// TIA Portal project "11_End_LAGER_Projekt_261019" (V17)

(* hardware
DEVICE "S7300/ET200M-Station_4"  S7-300 station
   slot 0: "Profilschiene_0"  Rail  6ES7 390-1***0-0AA0
   slot 1: "PS 307 5A_1"  PS 307 5A  6ES7 307-1EA01-0AA0
   slot 2: "PLC_WBS_Bus"  CPU 314C-2 DP  6ES7 314-6CH04-0AB0  V3.3
      slot 0: "MPI-Schnittstelle_1"  MPI
      slot 1: "DP-Schnittstelle_1"  DP
      slot 2: "DI 24/DO 16_1"  DI24/DO16
      slot 3: "AI 5/AO 2_1"  AI5/AO2
      slot 4: "Zählen_1"  Counter
      slot 5: "Positionieren_1"  Positioning
   slot 4: "DI 64x24VDC sinking/souring_1"  DI64 x 24VDC  6ES7 321-1BP00-0AA0
   slot 5: "DI 64x24VDC sinking/souring_2"  DI64 x 24VDC  6ES7 321-1BP00-0AA0
   slot 6: "DI 64x24VDC sinking/souring_3"  DI64 x 24VDC  6ES7 321-1BP00-0AA0
   slot 7: "DI 64x24VDC sinking/souring_4"  DI64 x 24VDC  6ES7 321-1BP00-0AA0
   slot 8: "DO 64x24VDC/0.3A sourcing_1"  DO64 x 24VDC / 0.3A, P  6ES7 322-1BP00-0AA0
   slot 9: "DO 64x24VDC/0.3A sourcing_2"  DO64 x 24VDC / 0.3A, P  6ES7 322-1BP00-0AA0
   slot 10: "DO 64x24VDC/0.3A sourcing_3"  DO64 x 24VDC / 0.3A, P  6ES7 322-1BP00-0AA0
   slot 11: "DO 64x24VDC/0.3A sourcing_4"  DO64 x 24VDC / 0.3A, P  6ES7 322-1BP00-0AA0
DEVICE "PC-System_1"  SIMATIC PC station
   slot 0: "SIMATIC PC-Station"  Rail  SIMATIC PC-Station  V1.0
      slot 125: "Stationmanager"  Station_Manager  V6.0.4
   slot 1: "HMI_RT_1"  WinCC RT Advanced  6AV2 104-0xxxx-xxxx  17.0.0.0
      slot 33792: "Computerschnittstelle"  Host interface
   slot 3: "CP 5711_1"  CP 5711  6GK1 571-1AA00  V7.1.1
*)

// ===== PLC "PLC_WBS_Bus"  CPU 314C-2 DP =====

VAR_GLOBAL   // PLC tag table "Standard-Variablentabelle"
   "test_taster" AT %M26.1 : Bool;
   "Tag_1" AT %M100.1 : Bool;
END_VAR

VAR_GLOBAL   // PLC tag table "Betriebsart"
   "S0_HS" AT %E0.0 : Bool;   // Hauptschalter 0-Aus, 1-Ein
   "S1_Not_Halt" AT %E0.1 : Bool;   // Not-Halt NC
   "S2_START" AT %E0.2 : Bool;   // Taster START NO
   "S3_STOP" AT %E0.3 : Bool;   // Taster STOP NC
   "Res_E06" AT %E0.6 : Bool;
   "Res_E07" AT %E0.7 : Bool;
   "Res_E10" AT %E1.0 : Bool;
   "Res_E11" AT %E1.1 : Bool;
   "Res_E12" AT %E1.2 : Bool;
   "Res_E13" AT %E1.3 : Bool;
   "Res_E14" AT %E1.4 : Bool;
   "Res_E15" AT %E1.5 : Bool;
   "Res_E16" AT %E1.6 : Bool;
   "Factory_IO_RUN" AT %E1.7 : Bool;   // Rückmeldung Factory IO läuft
   "P1_MS_RT" AT %A0.0 : Bool;   // Meldesäule Rot
   "P2_MS_GE" AT %A0.1 : Bool;   // Meldesäule Gelb
   "P3_MS_GN" AT %A0.2 : Bool;   // Meldesäule Grün
   "P10_START" AT %A0.3 : Bool;   // Anzeige grün in START-Taster
   "P11_STOP" AT %A0.4 : Bool;   // Anzeige gelb in START-Taster
   "Res_A0.5" AT %A0.5 : Bool;
   "P12_Anfahrwarnung" AT %A0.6 : Bool;   // Rundumleuchte System
   "P13_Sirene" AT %A0.7 : Bool;   // Sirene System
   "Res_A12" AT %A1.2 : Bool;
   "Res_A13" AT %A1.3 : Bool;
   "Res_A14" AT %A1.4 : Bool;
   "Res_A15" AT %A1.5 : Bool;
   "Res_A16" AT %A1.6 : Bool;
   "Res_A17" AT %A1.7 : Bool;
   "Log_1" AT %M0.1 : Bool;   // statisch "1"
   "Log_0" AT %M0.0 : Bool;   // statisch "0"
   "Takt_1HZ" AT %M100.5 : Bool;   // Taktmerker 1 Hz
   "Anzeige_Anzahl_Teile_BL" AT %AW22 : Int;   // Anzeige Teile blau im Lager
   "Anzeige_Anzahl_Teile_GN" AT %AW24 : Int;   // Anzeige Teile grün im Lager
   "Start_Merker" AT %M26.0 : Bool;
   "S4_Auswahl_GN" AT %E0.4 : Bool;   // Taster Auswahl Teile grün NO
   "S5_Auswahl_BL" AT %E0.5 : Bool;   // Taster Auswahl Teile blau NO
   "P14_Auswahl_GN" AT %A1.0 : Bool;   // Anzeige Auswahl grün Taster
   "P15_Auswahl_BL" AT %A1.1 : Bool;   // Anzeige Auswahl blau Taster
   "M_False" AT %M202.0 : Bool;
   "M_True" AT %M202.1 : Bool;
   "Takt_2,5Hz" AT %M100.2 : Bool;
   "Pult_EW" AT %EW0 : Word;
   "Pult_AW" AT %AW0 : Word;
END_VAR

VAR_GLOBAL   // PLC tag table "Lager"
   "B8001_RB8001" AT %E2.0 : Bool;   // Transportband-Anfang
   "B8802_RB8001" AT %E2.1 : Bool;   // Transportband-Ende
   "B8003_RB8002" AT %E2.2 : Bool;   // Transportband-Anfang
   "B8004_RB8002" AT %E2.3 : Bool;   // Transportband-Ende
   "B8005_RB8003" AT %E2.4 : Bool;   // Transportband-Anfang
   "B8006_RB8003" AT %E2.5 : Bool;   // Transportband-Ende
   "B8007_OT_BL" AT %E2.6 : Bool;
   "B8008_OT_GN" AT %E2.7 : Bool;
   "B8020_STAPL_8001_Endlage_links" AT %E3.0 : Bool;   // Regaltransportgerät
   "B8021_STAPL_8001_Mittel_Pos" AT %E3.1 : Bool;   // Regaltransportgerät
   "B8022_STAPL_8001_Endlage_rechts" AT %E3.2 : Bool;   // Regaltransportgerät
   "B8023_STAPL_Bew_X_aktiv" AT %E3.3 : Bool;   // Regaltransportgerät
   "B8024_STAPL_Bew_Z_aktiv" AT %E3.4 : Bool;   // Regaltransportgerät
   "Res_E35" AT %E3.5 : Bool;
   "Res_E36" AT %E3.6 : Bool;
   "Res_E37" AT %E3.7 : Bool;
   "RB8001" AT %A2.0 : Bool;
   "RB8002" AT %A2.1 : Bool;
   "RB8003" AT %A2.2 : Bool;
   "STAPL_8001_Palette_heben" AT %A2.3 : Bool;
   "STAPL_8001_links_ausfahren" AT %A2.4 : Bool;
   "STAPL_8001_rechts_ausfahren" AT %A2.5 : Bool;
   "P8001_Warnung_Bewegung_1" AT %A2.6 : Bool;   // Rundumleuchte
   "P8002_Warnung_Bewegung_2" AT %A2.7 : Bool;   // Rundumleuchte
   "Res_A30" AT %A3.0 : Bool;
   "Res_A31" AT %A3.1 : Bool;
   "Res_A32" AT %A3.2 : Bool;
   "Res_A33" AT %A3.3 : Bool;
   "Res_A34" AT %A3.4 : Bool;
   "Res_A35" AT %A3.5 : Bool;
   "Res_A36" AT %A3.6 : Bool;
   "Emitter_1" AT %A3.7 : Bool;   // Emitter_1
   "STAPL_8001_Fachposition" AT %AW20 : Int;
END_VAR

VAR_GLOBAL   // PLC tag table "Versand_1"
   "B9001_RB9001" AT %E4.0 : Bool;   // Transportband-Anfang
   "B9002_RB9001" AT %E4.1 : Bool;   // Transportband-Ende
   "B9003_RB9002" AT %E4.2 : Bool;   // Transportband-Anfang
   "B9004_RB9002" AT %E4.3 : Bool;   // Transportband-Ende
   "B9005_RB9003" AT %E4.4 : Bool;   // Transportband-Anfang
   "B9006_RB9003" AT %E4.5 : Bool;   // Transportband-Ende
   "B9007_OT_BL" AT %E4.6 : Bool;   // Farberkennung blau
   "B9008_OT_GN" AT %E4.7 : Bool;   // Farberkennung grün
   "B9020_STAPL_9001_Endlage_links" AT %E5.0 : Bool;   // Regaltransportgerät
   "B9021_STAPL_9001_Mittel_Pos" AT %E5.1 : Bool;   // Regaltransportgerät
   "B9022_STAPL_9001_Endlage_rechts" AT %E5.2 : Bool;   // Regaltransportgerät
   "B9023_STAPL_Bew_X_aktiv" AT %E5.3 : Bool;   // Regaltransportgerät
   "B9024_STAPL_Bew_Z_aktiv" AT %E5.4 : Bool;   // Regaltransportgerät
   "RB9001" AT %A4.0 : Bool;
   "RB9002" AT %A4.1 : Bool;
   "RB9003" AT %A4.2 : Bool;
   "STAPL_9001_Palette_heben" AT %A4.3 : Bool;
   "STAPL_9001_links_ausfahren" AT %A4.4 : Bool;
   "STAPL_9001_rechts_ausfahren" AT %A4.5 : Bool;
   "P9001_Warnung_Bewegung_1" AT %A4.6 : Bool;   // Rundumleuchte
   "P9002_Warnung_Bewegung_2" AT %A4.7 : Bool;   // Rundumleuchte
   "Res_A37" AT %A5.7 : Bool;
   "STAPL_9001_Fachposition" AT %AW26 : Int;
END_VAR

TYPE "Datenspeicher"
   STRUCT
      DatumUhrzeit : Date_And_Time;
      Materialfarbe : String[10];
      Materialfarbe_Nummer : Int;
      Frei : Bool := TRUE;
   END_STRUCT;
END_TYPE

TYPE "Pult_Output"
   STRUCT
      P1_MS_RT : Bool;
      P2_MS_GE : Bool;
      P3_MS_GN : Bool;
      P10_START : Bool;
      P11_STOP : Bool;
      "Res_A0.5" : Bool;
      P12_Anfahrwarnung : Bool;
      P13_Sirene : Bool;
      P14_Auswahl_GN : Bool;
      P15_Auswahl_BL : Bool;
      Res_A12 : Bool;
      Res_A13 : Bool;
      Res_A14 : Bool;
      Res_A15 : Bool;
      Res_A16 : Bool;
      Res_A17 : Bool;
   END_STRUCT;
END_TYPE

TYPE "Datenaustausch_Lager"
   STRUCT
      Anlage_Ein : Bool;
      Anlage_Betriebsbereit : Bool;
      Anlage_Stop : Bool;
      NotHalt : Bool;
      Position : Int;
   END_STRUCT;
END_TYPE

TYPE "Datenaustausch_Versand"
   STRUCT
      Anlage_Ein : Bool;
      Anlage_Betriebsbereit : Bool;
      Anlage_Stop : Bool;
      NotHalt : Bool;
      i_Blau : Bool;
      i_Grün : Bool;
      i_630_Grundstellung : Bool;
      i_640_RB_Frei : Bool;
      i_fehler : Bool;
      i_Blau_Anzahl : Int;
      i_Grün_Anzahl : Int;
      Position : Int;
   END_STRUCT;
END_TYPE

TYPE "Pult_Input"
   STRUCT
      S0_HS : Bool;
      S1_Not_Halt : Bool;
      S2_START : Bool;
      S3_STOP : Bool;
      S4_Auswahl_GN : Bool;
      S5_Auswahl_BL : Bool;
      Res_E06 : Bool;
      Res_E07 : Bool;
      Res_E10 : Bool;
      Res_E11 : Bool;
      Res_E12 : Bool;
      Res_E13 : Bool;
      Res_E14 : Bool;
      Res_E15 : Bool;
      Res_E16 : Bool;
      Factory_IO_RUN : Bool;
   END_STRUCT;
END_TYPE

// folder: LAGER/DB

DATA_BLOCK "HochregallagerDB"   // DB1
{ S7_Optimized_Access := 'FALSE' }
VERSION : 0.1
   VAR
      Freigabe : Bool := False;   // Freigabe der Anlage
      Palette_Bereit_Pos55 : Bool := True;   // Palette an Übergabeposition 55 zur Übernahme bereit
      Stapler_Fachposition_Eingabe : Int := 1;   // Zielposition des Staplers: 1–54 Lagerfach, 55 Übergabe
      Stapler_Auftrag_Aktiv : Bool;   // Stapler bearbeitet einen Auftrag
      Stapler_Auftrag_Fertig : Bool;   // Staplerauftrag abgeschlossen
      Stapler_Stoerung : Bool;   // Störung am Stapler vorhanden
      Farbe : Int;   // Erkannter Farbcode: 1 = Blau, 2 = Grün, 4 = Fehler
      Stappler_Aktuele_Farbe : Int;   // Farbcode der aktuell vom Stapler transportierten Palette
      Automatik : Bool := True;   // Automatikbetrieb aktiviert
      Motors_Ein : Bool;   // Einschaltsignal für die Rollenbahnmotoren
      Neue_Palette : Bool;   // Signal für eine neue Palette
      HMI_X_Bewegung : Int;   // Horizontale Position für die Stapleranimation im HMI
      HMI_Z_Bewegung : Int;   // Vertikale Position für die Stapleranimation im HMI
      Reset_Counter : Bool;   // Zähler zurücksetzen
      Lagerplaetze : Array[1..54] of "Datenspeicher";   // Lagerdaten der 54 Lagerplätze: Belegung, Farbe und Einlagerungszeit
      Anzahl_Blau : Int;   // Anzahl der eingelagerten blauen Paletten
      Anzahl_Gruen : Int;   // Anzahl der eingelagerten grünen Paletten
      Anzahl_Unbekannte_Farbe : Int;   // Anzahl der eingelagerten Unbekannte Paletten
      Einlagerungsposition : Int;   // Nummer des Lagerplatzes für die zu speichernden Palettendaten (1–54)
      Stapler_In_Bewegung : Bool;   // Stacker in motion
      Rollenbahn_In_Bewegung : Bool;   // Conveyor in motion
      Stoerung_Aktiv : Bool;   // Eine Störung liegt vor.
      Warnung_Aktiv : Bool;   // Eine Warnung liegt vor.
      Warnung_Wenig_Freie_Plaetze : Bool;   // TRUE: Warnschwelle erreicht oder unterschritten; auch bei vollem Lager aktiv.
      Lager_Voll : Bool;   // TRUE: Alle Lagerplaetze sind belegt.
      Stopp_Am_Zyklusende : Bool;
   END_VAR
BEGIN
END_DATA_BLOCK

DATA_BLOCK "HMI_Eingaben_DB"   // DB8
{ S7_Optimized_Access := 'FALSE' }
VERSION : 0.1
   VAR
      HMI_Start : Bool;
      HMI_Stop : Bool := TRUE;
      HMI_Not_Halt : Bool := TRUE;
      HMI_Hauptschalter : Bool;
      HMI_Start_Anzeige : Bool;
   END_VAR
BEGIN
END_DATA_BLOCK

// folder: LAGER/Instance

DATA_BLOCK "FB_Paketempfang_Rollenbahn_DB"   // DB2
{ S7_Optimized_Access := 'FALSE' }
VERSION : 0.1
// stored: InstanceOfName FB_Paketempfang_Rollenbahn
"FB_Paketempfang_Rollenbahn"
BEGIN
END_DATA_BLOCK

DATA_BLOCK "FB_Stapler_Ablauf_DB"   // DB3
{ S7_Optimized_Access := 'FALSE' }
VERSION : 0.1
// stored: InstanceOfName FB_Stapler_Ablauf
"FB_Stapler_Ablauf"
BEGIN
END_DATA_BLOCK

DATA_BLOCK "FB_Lagerverwaltung_DB"   // DB4
{ S7_Optimized_Access := 'FALSE' }
VERSION : 0.1
// stored: InstanceOfName FB_Lagerverwaltung
"FB_Lagerverwaltung"
BEGIN
END_DATA_BLOCK

DATA_BLOCK "FB_ControlPanel_DB"   // DB7
{ S7_Optimized_Access := 'FALSE' }
VERSION : 0.1
// stored: InstanceOfName FB_ControlPanel
"FB_ControlPanel"
BEGIN
END_DATA_BLOCK

DATA_BLOCK "Lager_Aufrufen_DB"   // DB9
{ S7_Optimized_Access := 'FALSE' }
VERSION : 0.1
// stored: InstanceOfName Lager_Aufrufen
"Lager_Aufrufen"
BEGIN
END_DATA_BLOCK

// folder: LAGER/Lager_AWL

DATA_BLOCK "Lager_Daten"   // DB8000
{ S7_Optimized_Access := 'FALSE' }
VERSION : 0.1
   VAR
      Lagerfach : Array[1..54] of Int;   // 1 = blau, 2 = grün, 0 = leer
   END_VAR
BEGIN
   Lagerfach[1] := 1;
   Lagerfach[2] := 2;
   Lagerfach[3] := 1;
   Lagerfach[4] := 2;
   Lagerfach[5] := 2;
   Lagerfach[6] := 2;
   Lagerfach[7] := 2;
   Lagerfach[8] := 2;
   Lagerfach[9] := 2;
   Lagerfach[10] := 2;
   Lagerfach[11] := 1;
   Lagerfach[12] := 1;
   Lagerfach[54] := 1;
   Lagerfach[13] := 1;
   Lagerfach[14] := 1;
   Lagerfach[15] := 1;
   Lagerfach[16] := 1;
   Lagerfach[17] := 1;
   Lagerfach[18] := 2;
   Lagerfach[19] := 2;
   Lagerfach[20] := 1;
   Lagerfach[21] := 2;
   Lagerfach[22] := 2;
   Lagerfach[23] := 2;
   Lagerfach[24] := 2;
   Lagerfach[25] := 2;
   Lagerfach[26] := 2;
   Lagerfach[27] := 2;
   Lagerfach[28] := 2;
   Lagerfach[29] := 1;
   Lagerfach[30] := 1;
   Lagerfach[31] := 1;
   Lagerfach[32] := 1;
   Lagerfach[33] := 1;
   Lagerfach[34] := 1;
   Lagerfach[35] := 1;
   Lagerfach[36] := 1;
   Lagerfach[37] := 1;
   Lagerfach[38] := 1;
   Lagerfach[39] := 2;
   Lagerfach[40] := 2;
   Lagerfach[41] := 2;
   Lagerfach[42] := 1;
   Lagerfach[43] := 1;
   Lagerfach[44] := 1;
   Lagerfach[45] := 1;
   Lagerfach[46] := 2;
   Lagerfach[47] := 2;
   Lagerfach[48] := 2;
   Lagerfach[49] := 2;
   Lagerfach[50] := 2;
   Lagerfach[51] := 0;
   Lagerfach[52] := 2;
   Lagerfach[53] := 1;
END_DATA_BLOCK

// folder: Versand

DATA_BLOCK "600_Versand_Main_DB"   // DB10
{ S7_Optimized_Access := 'FALSE' }
AUTHOR : DJonas
VERSION : 0.1
// stored: InstanceOfName 600_Versand_Main
"600_Versand_Main"
BEGIN
END_DATA_BLOCK

// folder: (top level)

ORGANIZATION_BLOCK "Main"   // OB1, FBD
TITLE = "Main Program Sweep (Cycle)"
{ S7_Optimized_Access := 'FALSE' }
VERSION : 0.1
   VAR_TEMP
      OB1_EV_CLASS : Byte;   // Bits 0-3 = 1 (Coming event), Bits 4-7 = 1 (Event class 1)
      OB1_SCAN_1 : Byte;   // 1 (Cold restart scan 1 of OB 1), 3 (Scan 2-n of OB 1)
      OB1_PRIORITY : Byte;   // Priority of OB Execution
      OB1_OB_NUMBR : Byte;   // 1 (Organization block 1, OB1)
      OB1_RESERVED_1 : Byte;   // Reserved for system
      OB1_RESERVED_2 : Byte;   // Reserved for system
      OB1_PREV_CYCLE : Int;   // Cycle time of previous OB1 scan (milliseconds)
      OB1_MIN_CYCLE : Int;   // Minimum cycle time of OB1 (milliseconds)
      OB1_MAX_CYCLE : Int;   // Maximum cycle time of OB1 (milliseconds)
      OB1_DATE_TIME : Date_And_Time;   // Date and time OB1 started
   END_VAR
BEGIN

REGION Network 1
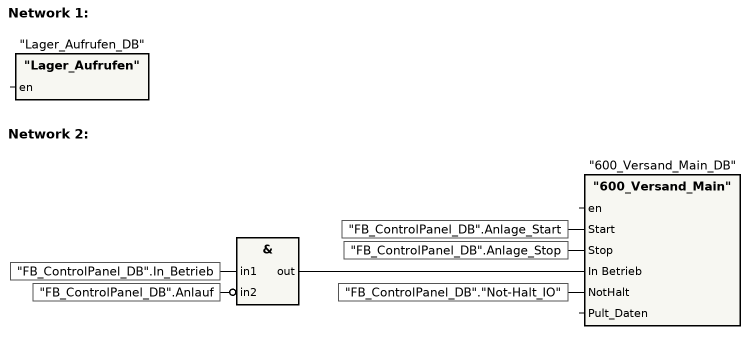
   "Lager_Aufrufen_DB"();   // "Lager_Aufrufen"
END_REGION

REGION Network 2
   "600_Versand_Main_DB"(Start := "FB_ControlPanel_DB".Anlage_Start,   // "600_Versand_Main"
                         Stop := "FB_ControlPanel_DB".Anlage_Stop,
                         "In Betrieb" := "FB_ControlPanel_DB".In_Betrieb AND NOT "FB_ControlPanel_DB".Anlauf,
                         NotHalt := "FB_ControlPanel_DB"."Not-Halt_IO");
END_REGION
END_ORGANIZATION_BLOCK

// folder: LAGER

FUNCTION_BLOCK "Lager_Aufrufen"   // FB4, FBD
{ S7_Optimized_Access := 'FALSE' }
VERSION : 0.1
BEGIN

REGION Network 1: Bedienpanel Signale verarbeiten
   // Start-, Stopp- und Not-Halt-Signale von Bedienpanel und HMI zusammenführen und an den FB_ControlPanel übergeben. Hauptschalter, Factory-I/O-Betriebsstatus und Palettenanzahlen einlesen sowie Meldeleuchten ansteuern.
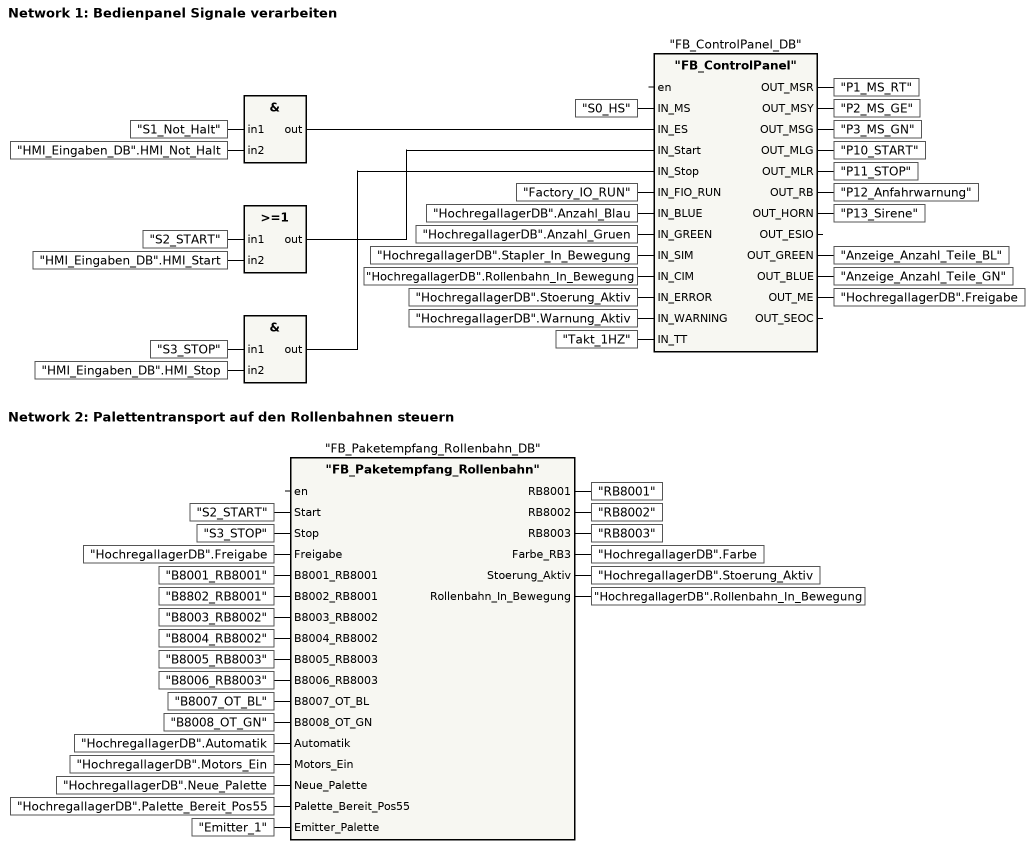
   "FB_ControlPanel_DB"(IN_MS := "S0_HS",   // "FB_ControlPanel"
                        IN_ES := "S1_Not_Halt" AND "HMI_Eingaben_DB".HMI_Not_Halt,
                        IN_Start := "S2_START" OR "HMI_Eingaben_DB".HMI_Start,
                        IN_Stop := "S3_STOP" AND "HMI_Eingaben_DB".HMI_Stop,
                        IN_FIO_RUN := "Factory_IO_RUN",
                        IN_BLUE := "HochregallagerDB".Anzahl_Blau,
                        IN_GREEN := "HochregallagerDB".Anzahl_Gruen,
                        IN_SIM := "HochregallagerDB".Stapler_In_Bewegung,
                        IN_CIM := "HochregallagerDB".Rollenbahn_In_Bewegung,
                        IN_ERROR := "HochregallagerDB".Stoerung_Aktiv,
                        IN_WARNING := "HochregallagerDB".Warnung_Aktiv,
                        IN_TT := "Takt_1HZ",
                        OUT_MSR => "P1_MS_RT",
                        OUT_MSY => "P2_MS_GE",
                        OUT_MSG => "P3_MS_GN",
                        OUT_MLG => "P10_START",
                        OUT_MLR => "P11_STOP",
                        OUT_RB => "P12_Anfahrwarnung",
                        OUT_HORN => "P13_Sirene",
                        OUT_GREEN => "Anzeige_Anzahl_Teile_BL",
                        OUT_BLUE => "Anzeige_Anzahl_Teile_GN",
                        OUT_ME => "HochregallagerDB".Freigabe);
END_REGION

REGION Network 2: Palettentransport auf den Rollenbahnen steuern
   // FB_Paketempfang_Rollenbahn aufrufen, Sensorsignale und Farberkennung auswerten sowie die drei Rollenbahnen abhängig von Start, Stopp und Freigabe ansteuern.
   "FB_Paketempfang_Rollenbahn_DB"(Start := "S2_START",   // "FB_Paketempfang_Rollenbahn"
                           Stop := "S3_STOP",
                           Freigabe := "HochregallagerDB".Freigabe,
                           B8001_RB8001 := "B8001_RB8001",
                           B8002_RB8001 := "B8802_RB8001",
                           B8003_RB8002 := "B8003_RB8002",
                           B8004_RB8002 := "B8004_RB8002",
                           B8005_RB8003 := "B8005_RB8003",
                           B8006_RB8003 := "B8006_RB8003",
                           B8007_OT_BL := "B8007_OT_BL",
                           B8008_OT_GN := "B8008_OT_GN",
                           Automatik := "HochregallagerDB".Automatik,
                           Motors_Ein := "HochregallagerDB".Motors_Ein,
                           Neue_Palette := "HochregallagerDB".Neue_Palette,
                           Palette_Bereit_Pos55 := "HochregallagerDB".Palette_Bereit_Pos55,
                           Emitter_Palette := "Emitter_1",
                           RB8001 => "RB8001",
                           RB8002 => "RB8002",
                           RB8003 => "RB8003",
                           Farbe_RB3 => "HochregallagerDB".Farbe,
                           Stoerung_Aktiv => "HochregallagerDB".Stoerung_Aktiv,
                           Rollenbahn_In_Bewegung => "HochregallagerDB".Rollenbahn_In_Bewegung);
END_REGION

REGION Network 3: Staplerablauf steuern
   // Der Baustein verarbeitet Freigabe, Stopp und Sensorsignale, steuert die Palettenaufnahme und Einlagerung und meldet den Auftragsstatus.
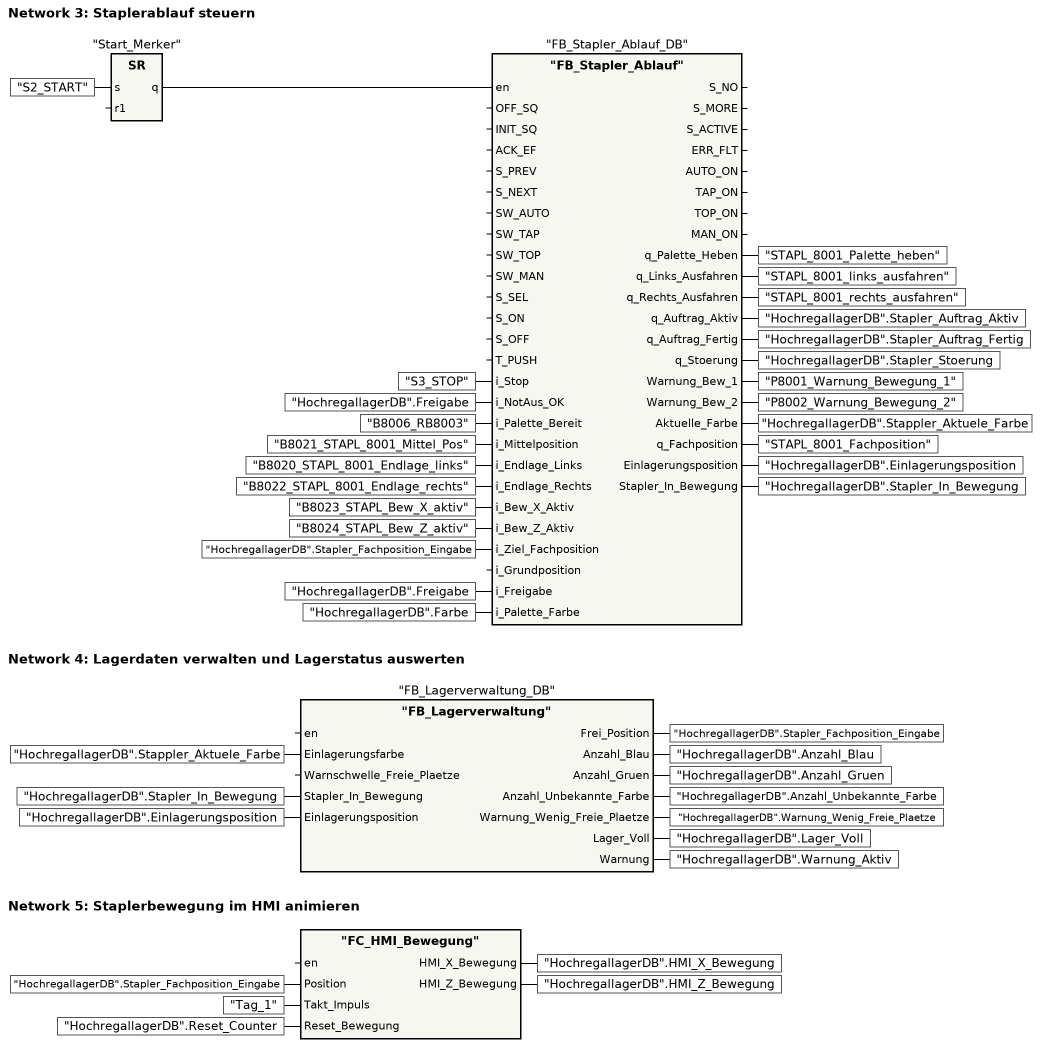
   IF "S2_START" THEN
       "Start_Merker" := TRUE;   // SR flip-flop
   END_IF;
   IF "Start_Merker" THEN
       "FB_Stapler_Ablauf_DB"(i_Stop := "S3_STOP",   // "FB_Stapler_Ablauf"
                              i_NotAus_OK := "HochregallagerDB".Freigabe,
                              i_Palette_Bereit := "B8006_RB8003",
                              i_Mittelposition := "B8021_STAPL_8001_Mittel_Pos",
                              i_Endlage_Links := "B8020_STAPL_8001_Endlage_links",
                              i_Endlage_Rechts := "B8022_STAPL_8001_Endlage_rechts",
                              i_Bew_X_Aktiv := "B8023_STAPL_Bew_X_aktiv",
                              i_Bew_Z_Aktiv := "B8024_STAPL_Bew_Z_aktiv",
                              i_Ziel_Fachposition := "HochregallagerDB".Stapler_Fachposition_Eingabe,
                              i_Freigabe := "HochregallagerDB".Freigabe,
                              i_Palette_Farbe := "HochregallagerDB".Farbe,
                              q_Palette_Heben => "STAPL_8001_Palette_heben",
                              q_Links_Ausfahren => "STAPL_8001_links_ausfahren",
                              q_Rechts_Ausfahren => "STAPL_8001_rechts_ausfahren",
                              q_Auftrag_Aktiv => "HochregallagerDB".Stapler_Auftrag_Aktiv,
                              q_Auftrag_Fertig => "HochregallagerDB".Stapler_Auftrag_Fertig,
                              q_Stoerung => "HochregallagerDB".Stapler_Stoerung,
                              Warnung_Bew_1 => "P8001_Warnung_Bewegung_1",
                              Warnung_Bew_2 => "P8002_Warnung_Bewegung_2",
                              Aktuelle_Farbe => "HochregallagerDB".Stappler_Aktuele_Farbe,
                              q_Fachposition => "STAPL_8001_Fachposition",
                              Einlagerungsposition => "HochregallagerDB".Einlagerungsposition,
                              Stapler_In_Bewegung => "HochregallagerDB".Stapler_In_Bewegung);
   END_IF;
END_REGION

REGION Network 4: Lagerdaten verwalten und Lagerstatus auswerten
   // FB_Lagerverwaltung aufrufen, Palettendaten speichern und freie Lagerplätze ermitteln. Paletten nach Farbe zählen und Warnungen bei wenigen freien Plätzen oder vollem Lager ausgeben.
   "FB_Lagerverwaltung_DB"(Einlagerungsfarbe := "HochregallagerDB".Stappler_Aktuele_Farbe,   // "FB_Lagerverwaltung"
                           Stapler_In_Bewegung := "HochregallagerDB".Stapler_In_Bewegung,
                           Einlagerungsposition := "HochregallagerDB".Einlagerungsposition,
                           Frei_Position => "HochregallagerDB".Stapler_Fachposition_Eingabe,
                           Anzahl_Blau => "HochregallagerDB".Anzahl_Blau,
                           Anzahl_Gruen => "HochregallagerDB".Anzahl_Gruen,
                           Anzahl_Unbekannte_Farbe => "HochregallagerDB".Anzahl_Unbekannte_Farbe,
                           Warnung_Wenig_Freie_Plaetze => "HochregallagerDB".Warnung_Wenig_Freie_Plaetze,
                           Lager_Voll => "HochregallagerDB".Lager_Voll,
                           Warnung => "HochregallagerDB".Warnung_Aktiv);
END_REGION

REGION Network 5: Staplerbewegung im HMI animieren
   // FC_HMI_Bewegung aufrufen, um aus der Fachposition und dem Taktsignal die X- und Z-Verschiebung für die HMI-Animation zu berechnen.
   "FC_HMI_Bewegung"(Position := "HochregallagerDB".Stapler_Fachposition_Eingabe,
                     Takt_Impuls := "Tag_1",
                     Reset_Bewegung := "HochregallagerDB".Reset_Counter,
                     HMI_X_Bewegung => "HochregallagerDB".HMI_X_Bewegung,
                     HMI_Z_Bewegung => "HochregallagerDB".HMI_Z_Bewegung);
END_REGION
END_FUNCTION_BLOCK

// folder: LAGER/FB

FUNCTION_BLOCK "FB_Paketempfang_Rollenbahn"   // FB1, FBD
TITLE = Paketempfang und Rollenbahnsteuerung
{ S7_Optimized_Access := 'FALSE' }
VERSION : 0.1
// - Der FB übernimmt die Steuerung des Palettentransports vom Emitter bis zur Übergabeposition 55 des Regalstapelsystems.
   VAR_INPUT
      Start : Bool;   // Anlage/Funktion freigegeben
      Stop : Bool;   // Stop-Anforderung
      Freigabe : Bool;   // Freigabe für Paketempfang und Rollenbahnsteuerung
      B8001_RB8001 : Bool;   // Sensor Palette auf Rollenbahn 1
      B8002_RB8001 : Bool;   // Sensor Ende Rollenbahn 1
      B8003_RB8002 : Bool;   // Sensor Palette auf Rollenbahn 2
      B8004_RB8002 : Bool;   // Sensor Ende Rollenbahn 2
      B8005_RB8003 : Bool;   // Sensor Palette auf Rollenbahn 3
      B8006_RB8003 : Bool;   // Sensor Ende Rollenbahn 3 (Palette hat Position 55 erreicht)
      B8007_OT_BL : Bool;   // optischer Sensor erkennt Blau
      B8008_OT_GN : Bool;   // optischer Sensor erkennt Grün
      Automatik : Bool;   // Betriebsart Automatik
      Motors_Ein : Bool;
      Neue_Palette : Bool;
   END_VAR
   VAR_OUTPUT
      RB8001 : Bool;   // Motor Rollenbahn 1
      RB8002 : Bool;   // Motor Rollenbahn 2
      RB8003 : Bool;   // Motor Rollenbahn 3
      Farbe_RB3 : Int;   // (1: Blau / 2:Grün / 4:Fehler)
      Stoerung_Aktiv : Bool;
      Rollenbahn_In_Bewegung : Bool;
   END_VAR
   VAR_IN_OUT
      Palette_Bereit_Pos55 : Bool;   // Palette steht zur Übernahme bereit
      Emitter_Palette : Bool;   // Emitter hat eine Palette bereitgestellt
   END_VAR
   VAR
      Empfang_Aktiv : Bool;   // FB bearbeitet aktuell eine Palette
      Betriebsfreigabe : Bool;   // Gespeicherte Freigabe für den Betrieb der Rollenbahnsteuerung
      Start_P_Merker : Bool;   // Flankenmerker für positive Flanke des Startsignals
      Emitter_P_Merker : Bool;   // Flankenmerker für positive Flanke des Emitter-Signals
      S2_N_Merker : Bool;   // Flankenmerker für negative Flanke von Sensor B8002
      S2_P_Merker : Bool;   // Merker für die positieve Flanke von Sensor 2
      S3_P_Merker : Bool;   // Flankenmerker für positive Flanke von Sensor B8003
      S4_N_Merker : Bool;   // Flankenmerker für negative Flanke von Sensor B8004
      S5_P_Merker : Bool;   // Flankenmerker für positive Flanke von Sensor B8005
      S6_N_Merker : Bool;   // Merker für die negative Flanke von Sensor 6
      S6_P_Merker : Bool;   // Flankenmerker für positive Flanke von Sensor B8006
      RB1_Merker : Bool;   // Speichermerker für Ansteuerung Rollenbahn 1
      RB2_Merker : Bool;   // Speichermerker für Ansteuerung Rollenbahn 2
      S3_N_Merker : Bool;
      RB3_Merker : Bool;   // Speichermerker für Ansteuerung Rollenbahn 3
      SBL_P_Merker : Bool;   // Flankenmerker für positive Flanke des Sensors Blau
      SGR_P_Merker : Bool;   // Flankenmerker für positive Flanke des Sensors Grün
      Palette_auf_RB1 : Bool;   // Palette befindet sich auf Rollenbahn 1
      Palette_auf_RB2 : Bool;   // Palette befindet sich auf Rollenbahn 2
      Palette_auf_RB3 : Bool;   // Palette befindet sich auf Rollenbahn 3
      Farbe_RB2 : Int;   // Erkannte Palettenfarbe auf Rollenbahn RB8002
      IEC_Timer_0_Instance : TON;   // Instanz des TON-Timers für Laufzeitüberwachung
      IEC_Timer_0_Instance_1 : TON;   // TON-Timerinstanz für Zeitüberwachung
      s_warnung_1 : Bool;   // Rollenbahn länger als zulässige Zeit aktiv
      s_warnung_2 : Bool;   // Sensor B8003_RB8002 länger als zulässige Zeit aktiv
      s_warnung_3 : Bool;
      IEC_Timer_0_Instance_2 : TON;
      Farbe_Merker : Bool;
      IEC_Timer_0_Instance_3 : TON;
   END_VAR
   VAR_TEMP   // added for the SCL form of the ladder/FBD networks
      _w1 : Bool;
      _w2 : Bool;
      _w3 : Bool;
      _w4 : Bool;
   END_VAR
BEGIN

REGION Network 1: Betriebsfreigabe
   // - Betriebsfreigabe über Start setzen und bei Stop bzw. fehlender Freigabe zurücksetzen.
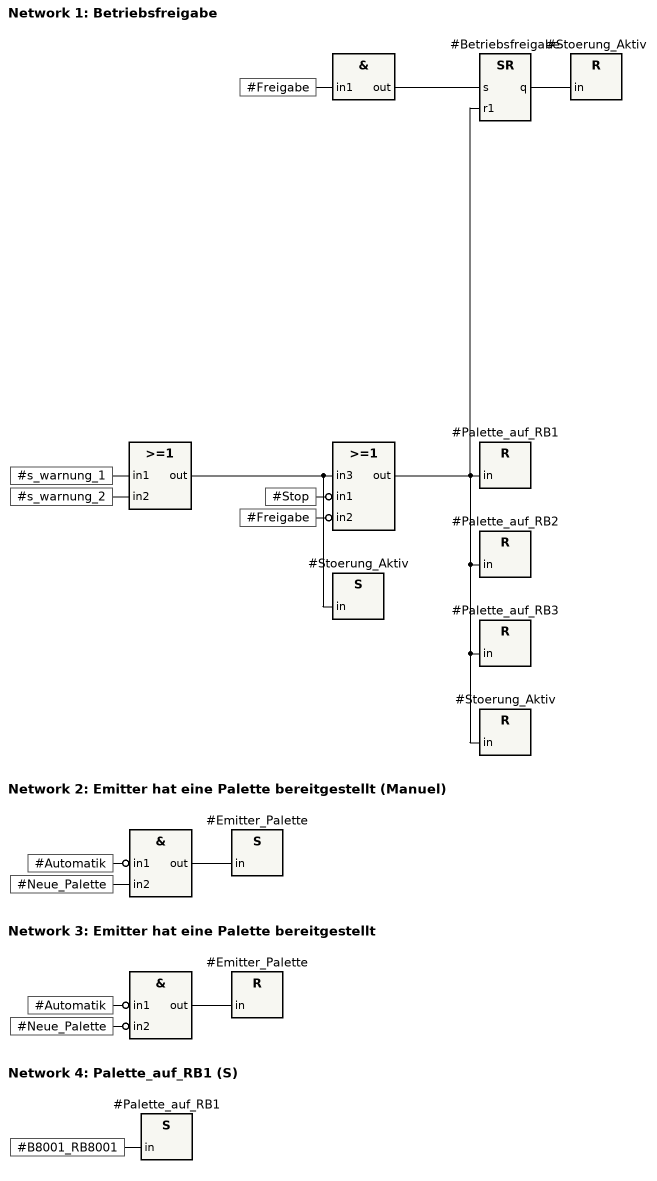
   #_w1 := #s_warnung_1 OR #s_warnung_2;
   #_w2 := #_w1 OR NOT #Stop OR NOT #Freigabe;
   IF #Freigabe THEN
       #Betriebsfreigabe := TRUE;   // SR flip-flop
   END_IF;
   IF #_w2 THEN #Betriebsfreigabe := FALSE; END_IF;
   IF #Betriebsfreigabe THEN #Stoerung_Aktiv := FALSE; END_IF;
   IF #_w2 THEN
       #Palette_auf_RB1 := FALSE;
       #Palette_auf_RB2 := FALSE;
       #Palette_auf_RB3 := FALSE;
       #Stoerung_Aktiv := FALSE;
   END_IF;
   IF #_w1 THEN #Stoerung_Aktiv := TRUE; END_IF;
END_REGION

REGION Network 2: Emitter hat eine Palette bereitgestellt (Manuel)
   IF NOT #Automatik AND #Neue_Palette THEN #Emitter_Palette := TRUE; END_IF;
END_REGION

REGION Network 3: Emitter hat eine Palette bereitgestellt
   IF NOT #Automatik AND NOT #Neue_Palette THEN #Emitter_Palette := FALSE; END_IF;
END_REGION

REGION Network 4: Palette_auf_RB1 (S)
   IF #B8001_RB8001 THEN #Palette_auf_RB1 := TRUE; END_IF;
END_REGION

REGION Network 5: Motor Rollenbahn 1
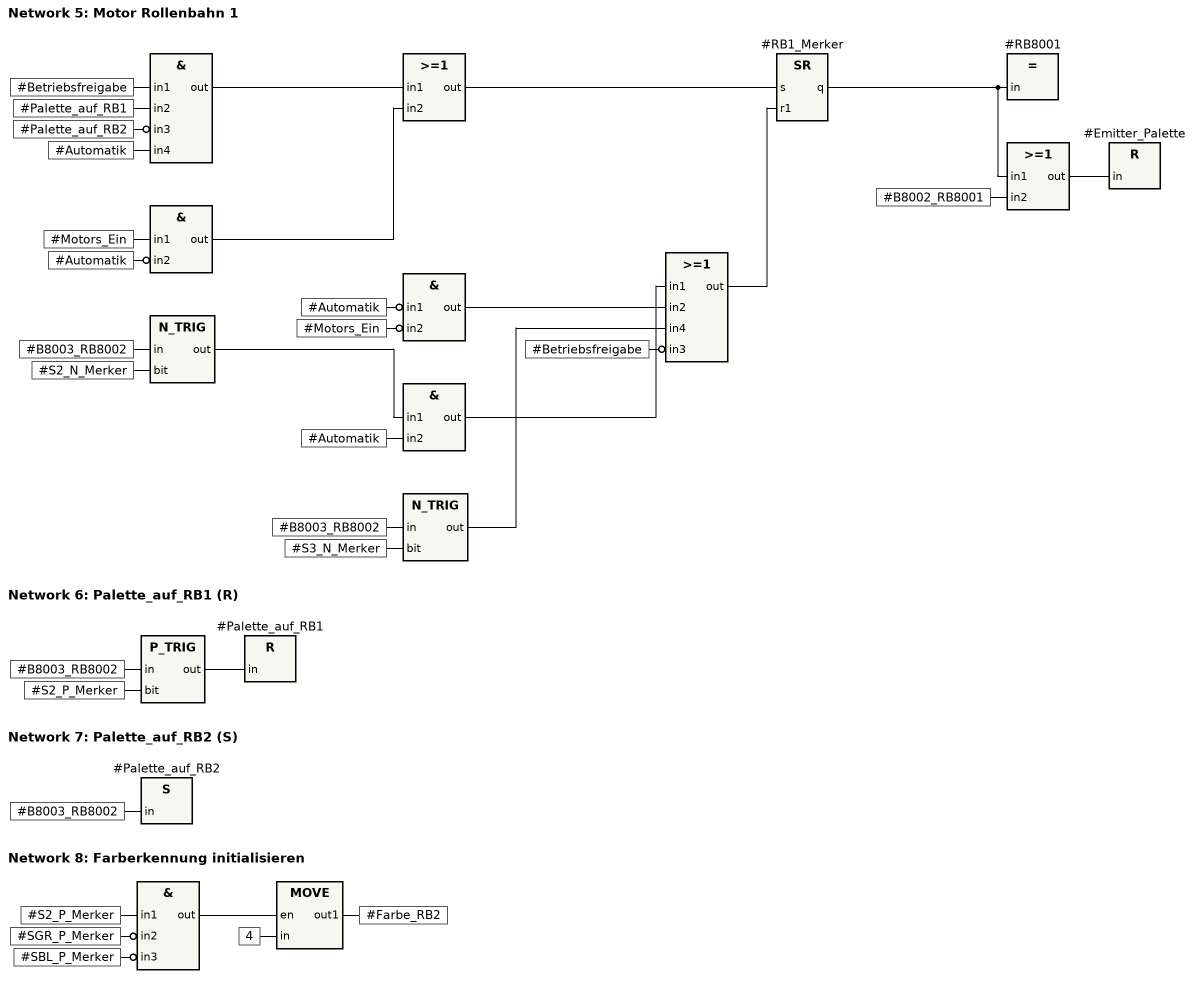
   #_w1 := NOT #B8003_RB8002 AND #S2_N_Merker;   // falling edge
   #S2_N_Merker := #B8003_RB8002;
   #_w2 := NOT #B8003_RB8002 AND #S3_N_Merker;   // falling edge
   #S3_N_Merker := #B8003_RB8002;
   IF (#Betriebsfreigabe AND #Palette_auf_RB1 AND NOT #Palette_auf_RB2 AND #Automatik) OR (#Motors_Ein AND NOT #Automatik) THEN
       #RB1_Merker := TRUE;   // SR flip-flop
   END_IF;
   IF (#_w1 AND #Automatik) OR (NOT #Automatik AND NOT #Motors_Ein) OR #_w2 OR NOT #Betriebsfreigabe THEN
       #RB1_Merker := FALSE;
   END_IF;
   #RB8001 := #RB1_Merker;
   IF #RB1_Merker OR #B8002_RB8001 THEN #Emitter_Palette := FALSE; END_IF;
END_REGION

REGION Network 6: Palette_auf_RB1 (R)
   #_w1 := #B8003_RB8002 AND NOT #S2_P_Merker;   // rising edge
   #S2_P_Merker := #B8003_RB8002;
   IF #_w1 THEN #Palette_auf_RB1 := FALSE; END_IF;
END_REGION

REGION Network 7: Palette_auf_RB2 (S)
   IF #B8003_RB8002 THEN #Palette_auf_RB2 := TRUE; END_IF;
END_REGION

REGION Network 8: Farberkennung initialisieren
   IF #S2_P_Merker AND NOT #SGR_P_Merker AND NOT #SBL_P_Merker THEN #Farbe_RB2 := 4; END_IF;
END_REGION

REGION Network 9: Motor Rollenbahn 2 / Farberkennung (Blau,Grün)
   // (1: Blau / 2:Grün / 4:Fehler)
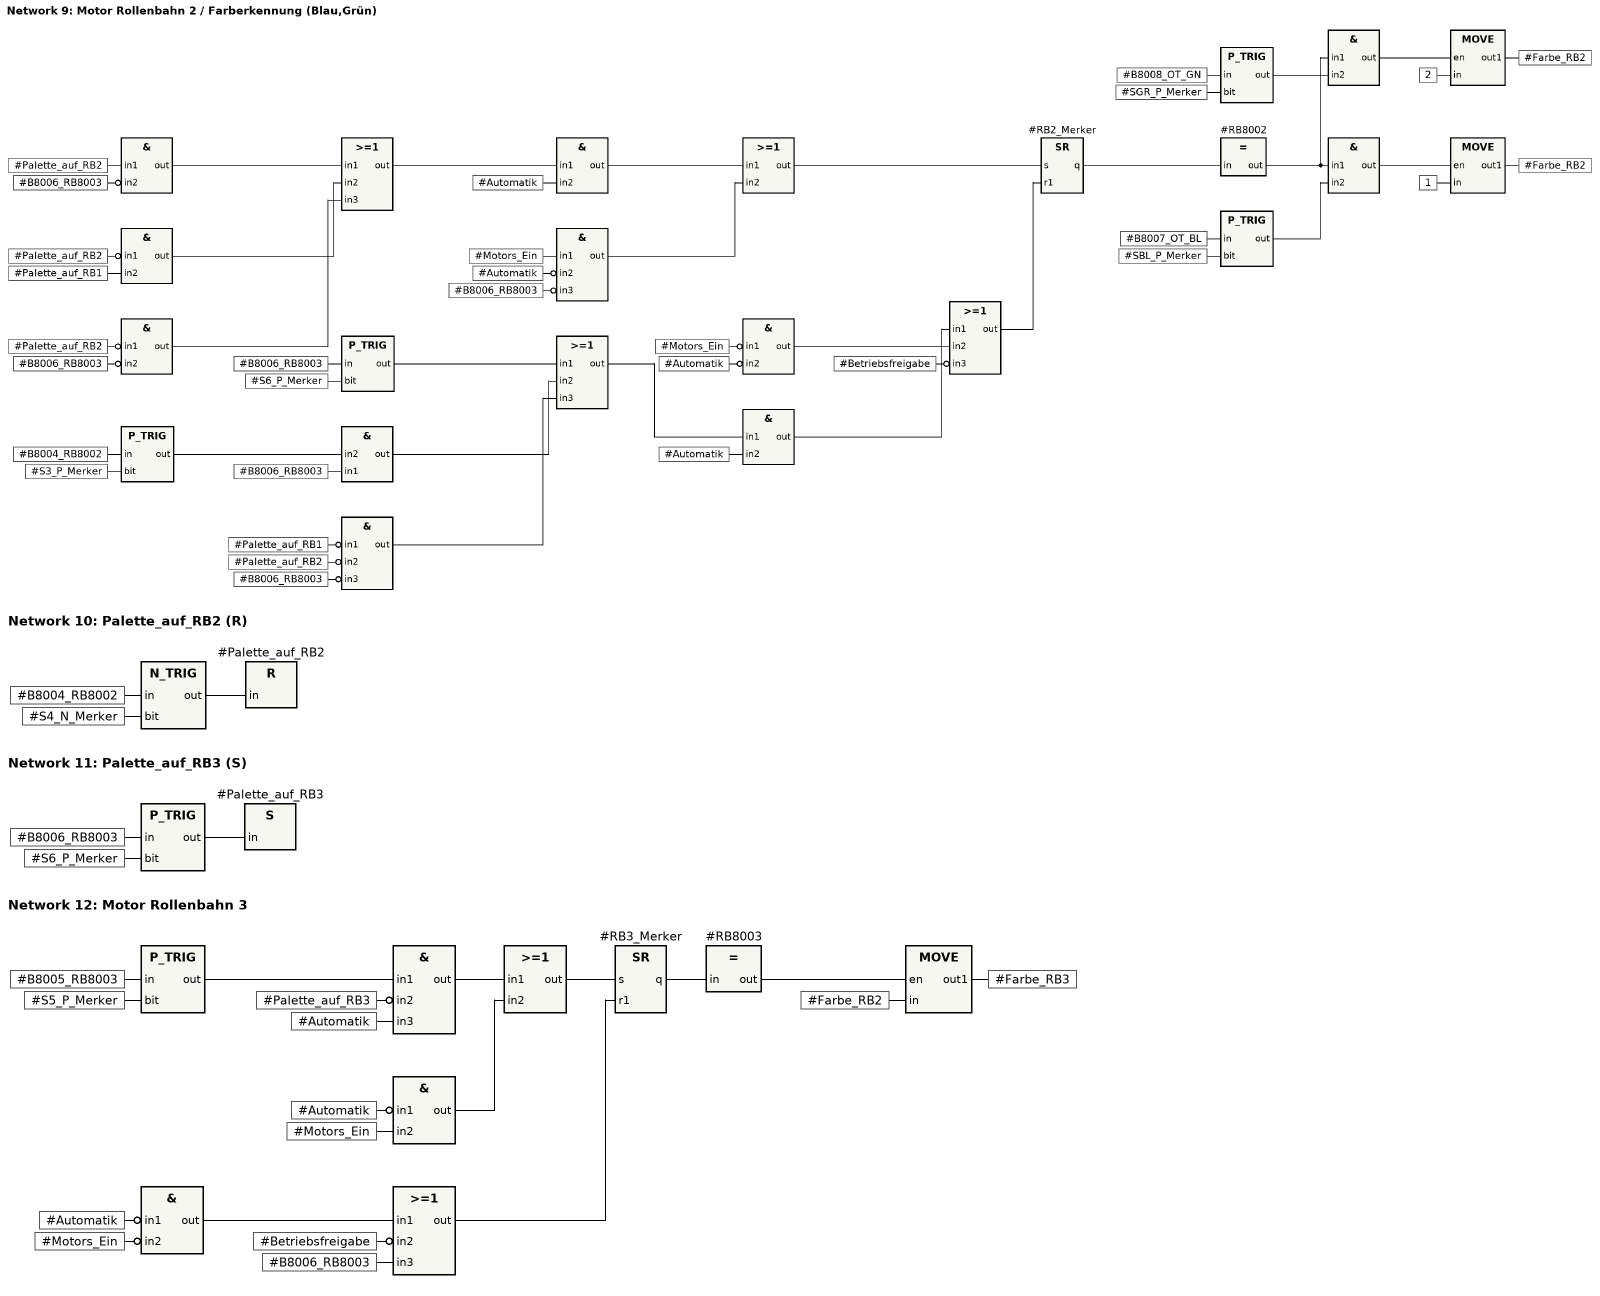
   #_w1 := #B8006_RB8003 AND NOT #S6_P_Merker;   // rising edge
   #S6_P_Merker := #B8006_RB8003;
   #_w2 := #B8004_RB8002 AND NOT #S3_P_Merker;   // rising edge
   #S3_P_Merker := #B8004_RB8002;
   IF (((#Palette_auf_RB2 AND NOT #B8006_RB8003) OR (NOT #Palette_auf_RB2 AND #Palette_auf_RB1) OR (NOT #Palette_auf_RB2 AND NOT #B8006_RB8003)) AND #Automatik) OR (#Motors_Ein AND NOT #Automatik AND NOT #B8006_RB8003) THEN
       #RB2_Merker := TRUE;   // SR flip-flop
   END_IF;
   IF ((#_w1 OR (#_w2 AND #B8006_RB8003) OR (NOT #Palette_auf_RB1 AND NOT #Palette_auf_RB2 AND NOT #B8006_RB8003)) AND #Automatik) OR (NOT #Motors_Ein AND NOT #Automatik) OR NOT #Betriebsfreigabe THEN
       #RB2_Merker := FALSE;
   END_IF;
   #RB8002 := #RB2_Merker;
   #_w3 := #B8008_OT_GN AND NOT #SGR_P_Merker;   // rising edge
   #SGR_P_Merker := #B8008_OT_GN;
   IF #RB2_Merker AND #_w3 THEN #Farbe_RB2 := 2; END_IF;
   #_w4 := #B8007_OT_BL AND NOT #SBL_P_Merker;   // rising edge
   #SBL_P_Merker := #B8007_OT_BL;
   IF #RB2_Merker AND #_w4 THEN #Farbe_RB2 := 1; END_IF;
END_REGION

REGION Network 10: Palette_auf_RB2 (R)
   #_w1 := NOT #B8004_RB8002 AND #S4_N_Merker;   // falling edge
   #S4_N_Merker := #B8004_RB8002;
   IF #_w1 THEN #Palette_auf_RB2 := FALSE; END_IF;
END_REGION

REGION Network 11: Palette_auf_RB3 (S)
   #_w1 := #B8006_RB8003 AND NOT #S6_P_Merker;   // rising edge
   #S6_P_Merker := #B8006_RB8003;
   IF #_w1 THEN #Palette_auf_RB3 := TRUE; END_IF;
END_REGION

REGION Network 12: Motor Rollenbahn 3
   // Farbe_RB3 (1: Blau / 2:Grün)
   #_w1 := #B8005_RB8003 AND NOT #S5_P_Merker;   // rising edge
   #S5_P_Merker := #B8005_RB8003;
   IF (#_w1 AND NOT #Palette_auf_RB3 AND #Automatik) OR (NOT #Automatik AND #Motors_Ein) THEN
       #RB3_Merker := TRUE;   // SR flip-flop
   END_IF;
   IF (NOT #Automatik AND NOT #Motors_Ein) OR NOT #Betriebsfreigabe OR #B8006_RB8003 THEN
       #RB3_Merker := FALSE;
   END_IF;
   #RB8003 := #RB3_Merker;
   IF #RB3_Merker THEN #Farbe_RB3 := #Farbe_RB2; END_IF;
END_REGION

REGION Network 13: Palette_auf_RB3 (R)
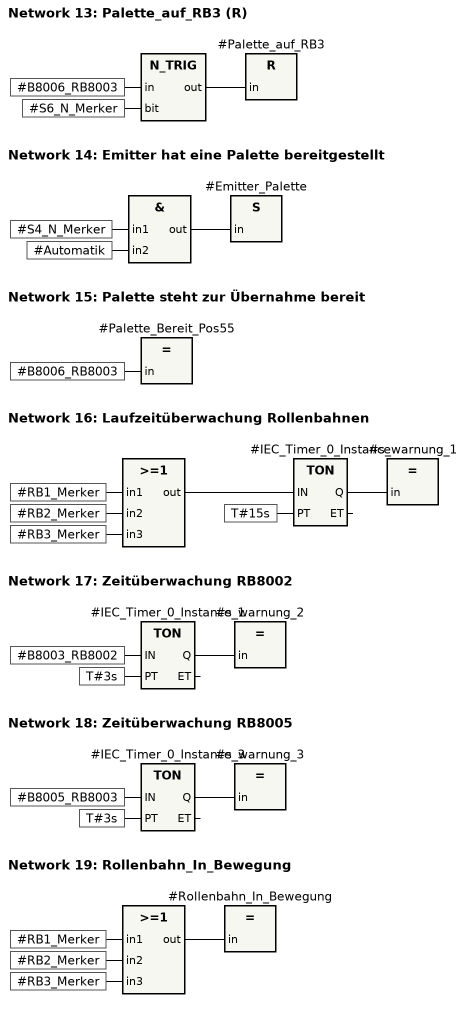
   #_w1 := NOT #B8006_RB8003 AND #S6_N_Merker;   // falling edge
   #S6_N_Merker := #B8006_RB8003;
   IF #_w1 THEN #Palette_auf_RB3 := FALSE; END_IF;
END_REGION

REGION Network 14: Emitter hat eine Palette bereitgestellt
   IF #S4_N_Merker AND #Automatik THEN #Emitter_Palette := TRUE; END_IF;
END_REGION

REGION Network 15: Palette steht zur Übernahme bereit
   #Palette_Bereit_Pos55 := #B8006_RB8003;
END_REGION

REGION Network 16: Laufzeitüberwachung Rollenbahnen
   // 14-s-Zeitüberwachung für aktive Rollenbahn. Bei Zeitüberschreitung wird s_warnung_1 gesetzt.
   #IEC_Timer_0_Instance.TON(IN := #RB1_Merker OR #RB2_Merker OR #RB3_Merker, PT := T#15s);
   #s_warnung_1 := #IEC_Timer_0_Instance.Q;
END_REGION

REGION Network 17: Zeitüberwachung RB8002
   // Ist der Sensor B8003_RB8002 länger als 4 s aktiv, wird die Warnung s_warnung_2 gesetzt.
   #IEC_Timer_0_Instance_1.TON(IN := #B8003_RB8002, PT := T#3s);
   #s_warnung_2 := #IEC_Timer_0_Instance_1.Q;
END_REGION

REGION Network 18: Zeitüberwachung RB8005
   #IEC_Timer_0_Instance_3.TON(IN := #B8005_RB8003, PT := T#3s);
   #s_warnung_3 := #IEC_Timer_0_Instance_3.Q;
END_REGION

REGION Network 19: Rollenbahn_In_Bewegung
   #Rollenbahn_In_Bewegung := #RB1_Merker OR #RB2_Merker OR #RB3_Merker;
END_REGION
END_FUNCTION_BLOCK

FUNCTION_BLOCK "FB_Stapler_Ablauf"   // FB2, GRAPH
{ S7_Optimized_Access := 'FALSE' }
VERSION : 0.1
   VAR_INPUT
      OFF_SQ : Bool := false;   // Kette ausschalten
      INIT_SQ : Bool := false;   // Kette in Initialzustand versetzen
      ACK_EF : Bool := false;   // Alle Fehler und Störungen quittieren
      S_PREV : Bool := false;   // Vorherigen Schritt am Parameter S_NO ausgeben
      S_NEXT : Bool := false;   // Nächsten Schritt am Parameter S_NO anzeigen
      SW_AUTO : Bool := false;   // Automatischer Betrieb
      SW_TAP : Bool := false;   // Halbautomatisch/Weiterschalten mit Transition
      SW_TOP : Bool := false;   // Halbautomatisch/Ignoriere Transition
      SW_MAN : Bool := false;   // Handbetrieb
      S_SEL : Int := 0;   // Schritt auswählen, der an S_NO ausgegeben werden soll
      S_ON : Bool := false;   // Schritt aktivieren, der an Parameter S_NO anliegt
      S_OFF : Bool := false;   // Schritt deaktivieren, der an Parameter S_NO anliegt
      T_PUSH : Bool := false;   // Schaltfreigabe für Transition im halbautomatischen Betrieb
      i_Stop : Bool;
      i_NotAus_OK : Bool;   // TRUE = kein Not-Aus / Anlage sicher
      i_Palette_Bereit : Bool;   // Palette wartet auf Einlagerung
      i_Mittelposition : Bool;   // Gabel in Mittelposition
      i_Endlage_Links : Bool;   // Gabel links vollständig ausgefahren
      i_Endlage_Rechts : Bool;   // Gabel rechts vollständig ausgefahren
      i_Bew_X_Aktiv : Bool;   // X-Bewegung aktiv
      i_Bew_Z_Aktiv : Bool;   // Z-Bewegung aktiv
      i_Ziel_Fachposition : Int;   // Zielposition für die Einlagerung
      i_Grundposition : Int := 55;   // Grundposition, bei dir 55
      i_Freigabe : Bool;
      i_Palette_Farbe : Int;   // (1: Blau / 2:Grün / 4:Fehler)
   END_VAR
   VAR_OUTPUT
      S_NO : Int := 0;   // Schrittnummer
      S_MORE : Bool := false;   // Weitere Schritte sind vorhanden und können in S_NO angezeigt werden.
      S_ACTIVE : Bool := false;   // Schritt, der an Parameter S_NO angezeigt wird, ist aktiv
      ERR_FLT : Bool := false;   // Sammelfehler Interlock oder Supervision
      AUTO_ON : Bool := false;   // Automatischer Betrieb eingeschaltet
      TAP_ON : Bool := false;   // Halbautomatischer Betrieb/Schritt mit Transition eingeschaltet
      TOP_ON : Bool := false;   // Halbautomatischer Betrieb/Ignoriere Transition eingeschaltet
      MAN_ON : Bool := false;   // Handbetrieb eingeschaltet
      q_Palette_Heben : Bool;   // Gabel links ausfahren
      q_Links_Ausfahren : Bool;   // Gabel links ausfahren
      q_Rechts_Ausfahren : Bool;   // Gabel rechts ausfahren
      q_Auftrag_Aktiv : Bool;   // Einlagerungsauftrag läuft
      q_Auftrag_Fertig : Bool;   // Auftrag abgeschlossen
      q_Stoerung : Bool;   // Störung im Staplerablauf
      Warnung_Bew_1 : Bool;
      Warnung_Bew_2 : Bool;
      Aktuelle_Farbe : Int;   // (1: Blau / 2:Grün / 4:Fehler)
      q_Fachposition : Int;   // Sollposition des Staplers
      Einlagerungsposition : Int;
      Stapler_In_Bewegung : Bool;
   END_VAR
   VAR
      SWITCH : Array[0..0] of DWord;
      SW_SQTS : Array[0..12] of Byte;
      SW_ADDR : Word := 16#1A;
      G7T_0 : GraphTransition;
      G7S_0 : GraphStep;
      PRE_CRIT : Array[0..0] of DWord;
      POST_CRIT : Array[0..0] of DWord;
      TVX : Array[0..2] of Byte;
      TTX : Array[0..2] of Byte;
      TSX : Array[0..2] of Byte;
      S00X : Array[0..2] of Byte;
      SOFFX : Array[0..2] of Byte;
      SONX : Array[0..2] of Byte;
      SAX : Array[0..2] of Byte;
      SERRX : Array[0..13] of Byte;
      SMX : Array[0..13] of Byte;
      S0X : Array[0..13] of Byte;
      S1X : Array[0..13] of Byte;
      S_DISPLAY : Int;   // Interne Anzeige des Ausgangsparameters S_NO
      S_SEL_OLD : Int;   // Vorheriger Wert an S_SEL
      S_DISPIDX : Byte;   // Index des Schritts, der an S_NO anliegt
      T_DISPIDX : Byte;   // Index der Transition, die an T_NO anliegt
      MOPEDGE : Struct
         AUTO : Bool := false;
         MAN : Bool := false;
         TAP : Bool := false;
         TOP : Bool := false;
         ACK_S : Bool := false;
         REG_S : Bool := false;
         T_PREV : Bool := false;
         T_NEXT : Bool := false;
         LOCK : Bool := false;
         SUP : Bool := false;
         ACKREQ : Bool := false;
         SSKIP : Bool := false;
         OFF : Bool := false;
         INIT : Bool := false;
         HALT : Bool := false;
         TMS_HALT : Bool := false;
         OPS_ZERO : Bool := false;
         SACT_DISP : Bool := false;
         SEF_DISP : Bool := false;
         SALL_DISP : Bool := false;
         S_PREV : Bool := false;
         S_NEXT : Bool := false;
         S_SELOK : Bool := false;
         S_ON : Bool := false;
         S_OFF : Bool := false;
         T_PUSH : Bool := false;
         REG : Bool := false;
         ACK : Bool := false;
         IL_PERM : Bool := false;
         T_PERM : Bool := false;
         ILP_MAN : Bool := false;
      END_STRUCT;
      MOP : Struct   // Betriebsart
         AUTO : Bool := true;   // Zustand: Automatischer Betrieb
         MAN : Bool := false;   // Zustand: Handbetrieb
         TAP : Bool := false;   // Zustand: Halbautomatisch/Weiterschalten mit Transition
         TOP : Bool := false;   // Zustand: Halbautomatisch/Ignoriere Transition
         ACK_S : Bool := false;   // Anforderung: Schritt quittieren, der an Parameter S_NO anliegt
         REG_S : Bool := false;   // Anforderung: Schritt registrieren, der an Parameter S_NO anliegt
         T_PREV : Bool := false;   // Anforderung: Vorherige gültige Transition am Parameter T_NO ausgeben
         T_NEXT : Bool := false;   // Anforderung: Nächste gültige Transition am Parameter T_NO ausgeben
         LOCK : Bool := true;   // Zustand: Interlockbearbeitung aktiviert
         SUP : Bool := true;   // Zustand: Supervisionsbearbeitung aktiviert
         ACKREQ : Bool := true;   // Zustand: Quittierung erforderlich
         SSKIP : Bool := false;   // Zustand: "Schritte überspringen" aktiviert
         OFF : Bool := false;   // Anforderung: Alle Schritte deaktivieren
         INIT : Bool := true;   // Anforderung: Kette in Initialzustand schalten
         HALT : Bool := false;   // Zustand: Kette schaltet nicht weiter
         TMS_HALT : Bool := false;   // Zustand: Alle internen Zeiten angehalten
         OPS_ZERO : Bool := false;   // Zustand: Alle mit N, L, D bearbeitete Operanden auf 0 gesetzt
         SACT_DISP : Bool := true;   // Zustand: Nur aktive Schritte anzeigen
         SEF_DISP : Bool := false;   // Zustand: Nur fehlerhafte und gestörte Schritte anzeigen
         SALL_DISP : Bool := false;   // Zustand: Alle Schritte anzeigen
         S_PREV : Bool := false;   // Anforderung: Vorherigen Schritt am Parameter S_NO ausgeben
         S_NEXT : Bool := false;   // Anforderung: Nächsten Schritt am Parameter S_NO ausgeben
         S_SELOK : Bool := false;   // Anforderung: Schrittnummer, die am Parameter S_SEL anliegt, am Parameter S_NO ausgeben
         S_ON : Bool := false;   // Anforderung: Schritt aktivieren, der am Parameter S_NO anliegt
         S_OFF : Bool := false;   // Anforderung: Schritt deaktivieren, der am Parameter S_NO anliegt
         T_PUSH : Bool := false;   // Anforderung: Schaltfreigabe für Transition
         REG : Bool := false;   // Anforderung: Alle Interlock- und Supervisionsfehler registrieren
         ACK : Bool := false;   // Anforderung: Alle Interlock- und Supervisionsfehler quittieren
         IL_PERM : Bool := false;   // Zustand: Permanente Bearbeitung aller Interlocks
         T_PERM : Bool := false;   // Zustand: Permanente Bearbeitung aller Transitionen
         ILP_MAN : Bool := false;   // Zustand: Permanente Bearbeitung aller Interlocks im Handbetrieb
      END_STRUCT;
      TICKS : Struct   // Zeittakte
         DELTA : Time := T#0ms;   // Zeitdifferenz zwischen zwei Zyklen
         OLD : Time := T#0ms;   // 10 ms Taktzählerstand im letzten Zyklus
         NEW : Time := T#0ms;   // 10 ms Taktzählerstand in diesem Zyklus
      END_STRUCT;
      SQ_FLAGS : Struct   // Kettenmerker
         ERR_FLT : Bool := false;   // Sammelfehler Interlock und Supervision
         ERROR : Bool := false;   // Sammelfehler Interlock
         FAULT : Bool := false;   // Sammelfehler Supervision
         RT_FAIL : Bool := false;   // Laufzeitfehler
         NO_SNO : Bool := false;   // Angeforderte Schrittnummer nicht gefunden
         NF_OFL : Bool := false;   // Überlauf: Zu viele Anforderungen ON oder OFF
         SA_OFL : Bool := false;   // Überlauf: Zu viele Schritte aktiv
         TV_OFL : Bool := false;   // Überlauf: Zu viele gültige Transitionen
         MSG_OFL : Bool := false;   // Überlauf: Nicht genügend Systemressourcen fü ALARM_S
         NO_SWI : Bool := false;   // Nicht Schalten in diesem Zyklus
         CYC_OP : Bool := false;   // Zyklische Bearbeitung der Kette nach Initialisierung
         AS_MSG : Bool := false;   // Meldungen zur Laufzeit durch Anweisung aktiviert oder deaktiviert
         AS_SEND : Bool := false;   // Meldungen von WR_USMSG senden oder nur in Diagnosepuffer eintragen
         SQ_BUSY : Bool := false;   // Interner Flankenmerker für Vorgangsbearbeitung
         SA_BUSY : Bool := false;   // Interner Flankenmerker für Vorgangsbearbeitung
         AS_SIG : Bool := false;   // Flankenmerker für Meldungen von Alarm_S und Alarm_SQ
      END_STRUCT;
      S_PTR : DWord := 16#7F0;
      S_PTR2 : DWord := 16#0;
      S_PTR3 : DWord := 16#1760;
      S_PTR4 : DWord := 16#16F0;
      T_PTR : DWord := 16#1680;
      C_AR2 : DWord := 16#0;
      M_FBDB : DWord := 16#20000;
      M_SNO : Word := 16#0;
      M_EVID : Word := 16#0;
      M_EVIL : DWord;
      M_EVSV : DWord;
      M_EV : DWord := 16#15B0;
      CRIT : Array[0..31] of Bool;
      S_START : Byte := 16#0;
      S_IDX : Byte := 16#0;
      S_INT : Int := 72;
      S_TMP : Byte := 16#0;
      T_START : Byte := 16#0;
      T_IDX : Byte := 16#0;
      T_TMP : Byte := 16#0;
      T_TMP2 : Byte := 16#00;
      TV_POT : Byte := 16#0E;
      RETURN1 : Byte := 16#0;
      RETURN2 : Byte := 16#0;
      SINI : Array[0..2] of Byte;
      LSTT : Array[0..12] of Byte;
      ATAJ : Array[0..12] of Byte;
      ATAB : Array[0..12] of Byte;
      PSTT : Array[0..12] of Byte;
      NSTT : Array[0..12] of Byte;
      ASSJ : Array[0..12] of Byte;
      ASSB : Array[0..12] of Byte;
      PTTS : Array[0..12] of Byte;
      NTTS : Array[0..12] of Byte;
      PRE_CNT : Word := 16#1;
      POST_CNT : Word := 16#1;
      ADR_COND : Word := 16#0;
      MAX_TVAL : Byte := 16#1;
      MAX_SACT : Byte := 16#1;
      MAX_CRIT : Byte := 16#4;
      T_CNT : Byte := 16#C;
      SUP_CNT : Byte := 16#0;
      LOCK_CNT : Byte := 16#2;
      S_CNT : Byte := 16#C;
      SQ_CNT : Byte := 16#1;
      PRS_INPAR : DWord := 16#E000FEC8;
      PRS_OUTPAR : DWord := 16#E000800F;
      GC_FLAGS : Struct
         T_MACH : Byte := 16#EB;
         COND_ED : Byte := 16#E2;
         W_LEVEL : Byte := 16#D5;
         FB_IF : Byte := 16#FA;
         AS_MSG : Word := 16#0;
         SSB : Word := 16#108;
         DILG : Word := 16#3FC;
         ADDR_T0 : Word := 16#2E;
         CRIT_AVAIL : Bool := false;
         SSKIP_AVAIL : Bool := true;
         SSKIP_ON : Bool := false;
         ACK_REQ : Bool := true;
         SYNC_AVAIL : Bool := true;
         ILP_MAN : Bool := false;
         SWM_LOCKED : Bool := false;
         SAVE_SW : Bool := true;
      END_STRUCT;
      G7_FBMARK : Byte := 16#3C;
      G7_RELEASE : Byte := 16#3C;
      G7_ID2 : Byte := 16#37;
      G7_ID1 : Byte := 16#47;
   END_VAR
   // SW_SQTS[0] := 16#1;
   // TVX[0] := 16#1;
   // TTX[0] := 16#1;
   // TSX[0] := 16#1;
   // S00X[0] := 16#1;
   // SOFFX[0] := 16#1;
   // SONX[0] := 16#1;
   // SAX[0] := 16#1;
   // SERRX[0] := 16#1;
   // SMX[0] := 16#1;
   // S0X[0] := 16#1;
   // S1X[0] := 16#1;
   // SINI[0] := 16#2;
   // SINI[1] := 16#1;
   // SINI[2] := 0;
   // LSTT[0] := 0;
   // LSTT[1] := 0;
   // LSTT[2] := 0;
   // LSTT[3] := 0;
   // LSTT[4] := 0;
   // LSTT[5] := 0;
   // LSTT[6] := 0;
   // LSTT[7] := 0;
   // ATAJ[0] := 0;
   // ATAJ[1] := 16#1;
   // ATAJ[2] := 16#2;
   // ATAJ[3] := 16#3;
   // ATAJ[4] := 16#4;
   // ATAJ[5] := 16#5;
   // ATAJ[6] := 16#6;
   // ATAJ[7] := 16#7;
   // ATAB[0] := 0;
   // ATAB[1] := 16#1;
   // ATAB[2] := 16#2;
   // ATAB[3] := 16#3;
   // ATAB[4] := 16#4;
   // ATAB[5] := 16#5;
   // ATAB[6] := 16#6;
   // ATAB[7] := 16#7;
   // PSTT[0] := 0;
   // PSTT[1] := 16#1;
   // PSTT[2] := 16#2;
   // PSTT[3] := 16#3;
   // PSTT[4] := 16#4;
   // PSTT[5] := 16#5;
   // PSTT[6] := 16#6;
   // PSTT[7] := 16#7;
   // NSTT[0] := 16#1;
   // NSTT[1] := 16#2;
   // NSTT[2] := 16#3;
   // NSTT[3] := 16#4;
   // NSTT[4] := 16#5;
   // NSTT[5] := 16#6;
   // NSTT[6] := 16#7;
   // NSTT[7] := 16#8;
   // ASSJ[0] := 0;
   // ASSJ[1] := 16#1;
   // ASSJ[2] := 16#2;
   // ASSJ[3] := 16#3;
   // ASSJ[4] := 16#4;
   // ASSJ[5] := 16#5;
   // ASSJ[6] := 16#6;
   // ASSJ[7] := 16#7;
   // ASSB[0] := 0;
   // ASSB[1] := 16#1;
   // ASSB[2] := 16#2;
   // ASSB[3] := 16#3;
   // ASSB[4] := 16#4;
   // ASSB[5] := 16#5;
   // ASSB[6] := 16#6;
   // ASSB[7] := 16#7;
   // PTTS[0] := 0;
   // PTTS[2] := 16#1;
   // PTTS[3] := 16#2;
   // PTTS[4] := 16#3;
   // PTTS[5] := 16#4;
   // PTTS[6] := 16#5;
   // PTTS[7] := 16#6;
   // NTTS[0] := 0;
   // NTTS[1] := 16#1;
   // NTTS[2] := 16#2;
   // NTTS[3] := 16#3;
   // NTTS[4] := 16#4;
   // NTTS[5] := 16#5;
   // NTTS[6] := 16#6;
   // NTTS[7] := 16#7;
   // LSTT[8] := 0;
   // LSTT[9] := 0;
   // LSTT[10] := 0;
   // ATAJ[8] := 16#8;
   // ATAJ[9] := 16#9;
   // ATAJ[10] := 16#A;
   // ATAB[8] := 16#8;
   // ATAB[9] := 16#9;
   // ATAB[10] := 16#A;
   // PSTT[8] := 16#8;
   // PSTT[9] := 16#9;
   // PSTT[10] := 16#A;
   // NSTT[8] := 16#9;
   // NSTT[9] := 16#A;
   // NSTT[10] := 16#C;
   // ASSJ[8] := 16#8;
   // ASSJ[9] := 16#9;
   // ASSJ[10] := 16#A;
   // ASSB[8] := 16#8;
   // ASSB[9] := 16#9;
   // ASSB[10] := 16#A;
   // PTTS[8] := 16#7;
   // PTTS[9] := 16#8;
   // PTTS[10] := 16#9;
   // NTTS[8] := 16#8;
   // NTTS[9] := 16#9;
   // NTTS[10] := 16#A;
   // LSTT[11] := 16#1;
   // ATAJ[11] := 16#B;
   // ATAB[11] := 16#B;
   // PSTT[11] := 16#B;
   // NSTT[11] := 16#1;
   // ASSJ[11] := 16#B;
   // ASSB[11] := 16#B;
   // PTTS[11] := 16#C;
   // NTTS[11] := 16#B;
   // LSTT[12] := 0;
   // ATAJ[12] := 16#C;
   // ATAB[12] := 16#C;
   // PSTT[12] := 16#C;
   // NSTT[12] := 16#B;
   // ASSJ[12] := 16#C;
   // ASSB[12] := 16#C;
   // PTTS[12] := 16#A;
   // NTTS[12] := 16#C;
BEGIN
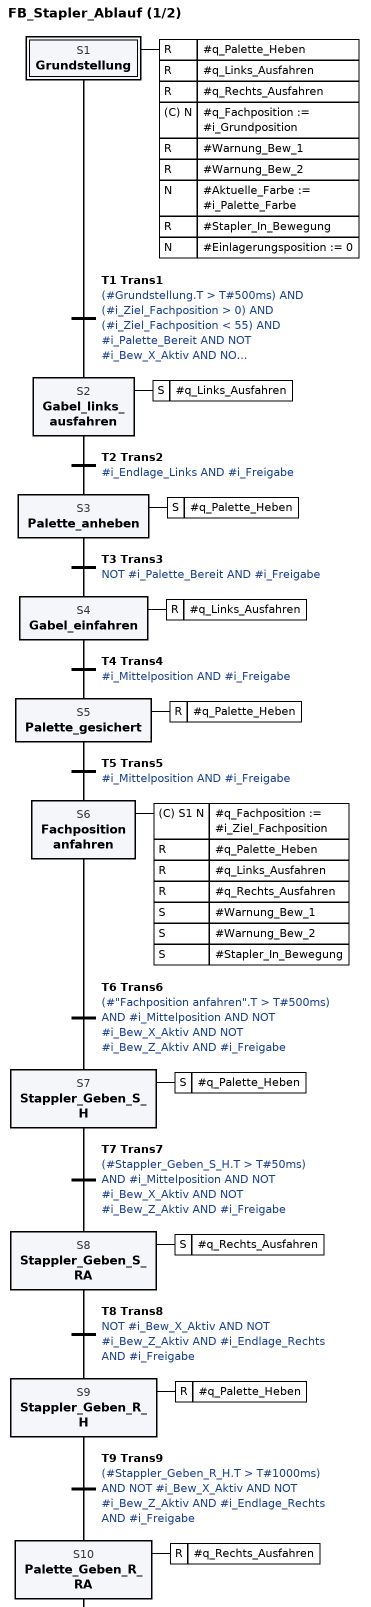
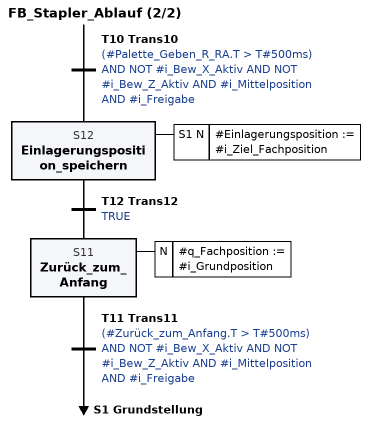
   // sequencer 1
   INITIAL_STEP Grundstellung:   // S1
      interlock C := #i_NotAus_OK AND #i_Stop;
      // - Stapler befindet sich in Grundstellung auf Position 55. Alle Ausgänge sind deaktiviert. Warten auf eine einlagerbereite Palette.
              R    #q_Palette_Heben
              R    #q_Links_Ausfahren
              R    #q_Rechts_Ausfahren
      (C)     N    #q_Fachposition := #i_Grundposition
              R    #Warnung_Bew_1
              R    #Warnung_Bew_2
              N    #Aktuelle_Farbe := #i_Palette_Farbe
              R    #Stapler_In_Bewegung
              N    #Einlagerungsposition := 0
   END_STEP
   TRANSITION Trans1 FROM Grundstellung TO Gabel_links_ausfahren   // T1
      := (#Grundstellung.T > T#500ms) AND (#i_Ziel_Fachposition > 0) AND (#i_Ziel_Fachposition < 55) AND #i_Palette_Bereit AND NOT #i_Bew_X_Aktiv AND NOT #i_Bew_Z_Aktiv AND #i_NotAus_OK AND #i_Stop AND #i_Freigabe;
   END_TRANSITION
   STEP Gabel_links_ausfahren:   // S2
              S    #q_Links_Ausfahren
   END_STEP
   TRANSITION Trans2 FROM Gabel_links_ausfahren TO Palette_anheben   // T2
      := #i_Endlage_Links AND #i_Freigabe;
   END_TRANSITION
   STEP Palette_anheben:   // S3
              S    #q_Palette_Heben
   END_STEP
   TRANSITION Trans3 FROM Palette_anheben TO Gabel_einfahren   // T3
      := NOT #i_Palette_Bereit AND #i_Freigabe;
   END_TRANSITION
   STEP Gabel_einfahren:   // S4
              R    #q_Links_Ausfahren
   END_STEP
   TRANSITION Trans4 FROM Gabel_einfahren TO Palette_gesichert   // T4
      := #i_Mittelposition AND #i_Freigabe;
   END_TRANSITION
   STEP Palette_gesichert:   // S5
              R    #q_Palette_Heben
   END_STEP
   TRANSITION Trans5 FROM Palette_gesichert TO "Fachposition anfahren"   // T5
      := #i_Mittelposition AND #i_Freigabe;
   END_TRANSITION
   STEP "Fachposition anfahren":   // S6
      interlock C := #i_Freigabe;
      // - Bei erfülltem Interlock wird die Ziel-Fachposition an den Stapler übergeben. - Die Ausgänge für Palette heben sowie Gabel links/rechts ausfahren werden zurückgesetzt. - Die Bewegungswarnungen werden gesetzt.
      (C) S1  N    #q_Fachposition := #i_Ziel_Fachposition
              R    #q_Palette_Heben
              R    #q_Links_Ausfahren
              R    #q_Rechts_Ausfahren
              S    #Warnung_Bew_1
              S    #Warnung_Bew_2
              S    #Stapler_In_Bewegung
   END_STEP
   TRANSITION Trans6 FROM "Fachposition anfahren" TO Stappler_Geben_S_H   // T6
      := (#"Fachposition anfahren".T > T#500ms) AND #i_Mittelposition AND NOT #i_Bew_X_Aktiv AND NOT #i_Bew_Z_Aktiv AND #i_Freigabe;
   END_TRANSITION
   STEP Stappler_Geben_S_H:   // S7
              S    #q_Palette_Heben
   END_STEP
   TRANSITION Trans7 FROM Stappler_Geben_S_H TO Stappler_Geben_S_RA   // T7
      := (#Stappler_Geben_S_H.T > T#50ms) AND #i_Mittelposition AND NOT #i_Bew_X_Aktiv AND NOT #i_Bew_Z_Aktiv AND #i_Freigabe;
   END_TRANSITION
   STEP Stappler_Geben_S_RA:   // S8
              S    #q_Rechts_Ausfahren
   END_STEP
   TRANSITION Trans8 FROM Stappler_Geben_S_RA TO Stappler_Geben_R_H   // T8
      := NOT #i_Bew_X_Aktiv AND NOT #i_Bew_Z_Aktiv AND #i_Endlage_Rechts AND #i_Freigabe;
   END_TRANSITION
   STEP Stappler_Geben_R_H:   // S9
              R    #q_Palette_Heben
   END_STEP
   TRANSITION Trans9 FROM Stappler_Geben_R_H TO Palette_Geben_R_RA   // T9
      := (#Stappler_Geben_R_H.T > T#1000ms) AND NOT #i_Bew_X_Aktiv AND NOT #i_Bew_Z_Aktiv AND #i_Endlage_Rechts AND #i_Freigabe;
   END_TRANSITION
   STEP Palette_Geben_R_RA:   // S10
              R    #q_Rechts_Ausfahren
   END_STEP
   TRANSITION Trans10 FROM Palette_Geben_R_RA TO Einlagerungsposition_speichern   // T10
      := (#Palette_Geben_R_RA.T > T#500ms) AND NOT #i_Bew_X_Aktiv AND NOT #i_Bew_Z_Aktiv AND #i_Mittelposition AND #i_Freigabe;
   END_TRANSITION
   STEP Zurück_zum_Anfang:   // S11
              N    #q_Fachposition := #i_Grundposition
   END_STEP
   TRANSITION Trans11 FROM Zurück_zum_Anfang TO Grundstellung   // T11, jump
      := (#Zurück_zum_Anfang.T > T#500ms) AND NOT #i_Bew_X_Aktiv AND NOT #i_Bew_Z_Aktiv AND #i_Mittelposition AND #i_Freigabe;
   END_TRANSITION
   STEP Einlagerungsposition_speichern:   // S12
      // - Beim Aktivieren des Schrittes wird die Ziel-Fachposition als Einlagerungsposition gespeichert. - Der FB_Lagerverwaltung verwendet diese Position, um die Palettendaten im Lagerarray zu speichern und anschließend den nächsten freien Lagerplatz zu ermitteln.
          S1  N    #Einlagerungsposition := #i_Ziel_Fachposition
   END_STEP
   TRANSITION Trans12 FROM Einlagerungsposition_speichern TO Zurück_zum_Anfang   // T12
      := TRUE;
   END_TRANSITION
END_FUNCTION_BLOCK

FUNCTION_BLOCK "FB_Lagerverwaltung"   // FB3, SCL
{ S7_Optimized_Access := 'FALSE' }
VERSION : 0.1
   VAR_INPUT
      Einlagerungsfarbe : Int;   // Farbcode der einzulagernden Palette: 1 = Blau, 2 = Gruen, 4 = Fehler
      Warnschwelle_Freie_Plaetze : Int := 5;   // Warnung bei dieser Anzahl freier Lagerplaetze oder weniger.
      Stapler_In_Bewegung : Bool;
   END_VAR
   VAR_OUTPUT
      Frei_Position : Int := 1;   // Kleinste freie Lagerplatznummer (1–54); 0 = kein freier Lagerplatz.
      Anzahl_Blau : Int;   // Anzahl der eingelagerten blauen Paletten.
      Anzahl_Gruen : Int;   // Anzahl der eingelagerten gruenen Paletten.
      Anzahl_Unbekannte_Farbe : Int;
      Warnung_Wenig_Freie_Plaetze : Bool;   // Warnschwelle erreicht: Nur noch wenige freie Lagerplätze verfügbar.
      Lager_Voll : Bool;   // TRUE: Alle Lagerplaetze sind belegt.
      Warnung : Bool;   // Sammelwarnung: Wenige freie Lagerplaetze oder Lager voll.
   END_VAR
   VAR_IN_OUT
      Einlagerungsposition : Int;   // Ziellagerplatz zum Speichern der Palettendaten (1–54).
   END_VAR
   VAR
      Einlagerungszeit : Date_And_Time;   // Von der CPU gelesener Zeitstempel der Einlagerung.
      Status_Uhrzeit : Int;   // Rueckgabecode von RD_SYS_T: 0 = erfolgreich, sonst Fehler.
      i : Int := 1;   // Schleifenindex zum Durchlaufen der 54 Lagerplaetze.
   END_VAR
   VAR_TEMP
      Anzahl_Freie_Plaetze : Int;   // Aktuelle Anzahl der freien Lagerplaetze (0–54).
   END_VAR
BEGIN
   // =====================================================
   // 1. Gueltigkeit der Einlagerungsposition pruefen
   // Nur Lagerplaetze von 1 bis 54 sind zulaessig.
   // =====================================================
   REGION Palettendaten speichern und Lagerplatz belegen

       IF (#Einlagerungsposition >= 1) AND (#Einlagerungsposition <= 54) THEN
           // =================================================
           // 1. Belegungsstatus pruefen
           // Daten nur in einen freien Lagerplatz schreiben.
           // Vorhandene Daten belegter Plaetze bleiben erhalten.
           // =================================================
           IF "HochregallagerDB".Lagerplaetze[#Einlagerungsposition].Frei THEN

               // =============================================
               // 2. Aktuelles Datum und Uhrzeit der CPU lesen
               // Status_Uhrzeit enthaelt den Rueckgabecode.
               // 0 = Zeit erfolgreich gelesen.
               // =============================================
               #Status_Uhrzeit := RD_SYS_T(OUT => #Einlagerungszeit);

               // =============================================
               // 3. Zeitstempel und numerischen Farbcode speichern
               // 1 = Blau, 2 = Gruen, 4 = Fehler.
               // =============================================
               "HochregallagerDB".Lagerplaetze[#Einlagerungsposition].DatumUhrzeit :=
               #Einlagerungszeit;

               "HochregallagerDB".Lagerplaetze[#Einlagerungsposition].Materialfarbe_Nummer :=
               #Einlagerungsfarbe;

               // =============================================
               // 4. Farbcode in einen lesbaren Text umwandeln
               // Nicht definierte Farbcodes werden als
               // 'Unbekannt' gespeichert.
               // =============================================
               CASE #Einlagerungsfarbe OF
                   1:
                       "HochregallagerDB".Lagerplaetze[#Einlagerungsposition].Materialfarbe :=
                       'Blau';
                   2:
                       "HochregallagerDB".Lagerplaetze[#Einlagerungsposition].Materialfarbe :=
                       'Gruen';
                   4:
                       "HochregallagerDB".Lagerplaetze[#Einlagerungsposition].Materialfarbe :=
                       'Fehler';
                   ELSE
                       "HochregallagerDB".Lagerplaetze[#Einlagerungsposition].Materialfarbe :=
                       'Unbekannt';
               END_CASE;

               // =============================================
               // 5. Lagerplatz als belegt markieren
               // Frei = FALSE: belegt; Frei = TRUE: frei.
               // =============================================
               "HochregallagerDB".Lagerplaetze[#Einlagerungsposition].Frei :=
               FALSE;

               #Einlagerungsposition := 0;
           END_IF;

       END_IF;
   END_REGION

   // =====================================================
   // 2. Kleinsten freien Lagerplatz ermitteln
   // Aufsteigende Suche von Platz 1 bis 54.
   // Beim ersten freien Platz wird die Suche beendet.
   // Frei_Position = 0 bedeutet: kein freier Platz vorhanden.
   // =====================================================
   REGION Freien Lagerplatz suchen
       IF NOT #Stapler_In_Bewegung THEN
           #Frei_Position := 0;
           FOR #i := 1 TO 54 DO
               IF "HochregallagerDB".Lagerplaetze[#i].Frei THEN
                   #Frei_Position := #i;
                   EXIT;
               END_IF;
           END_FOR;
           ;
       END_IF;
   END_REGION

   // =====================================================
   // 3. Blaue und gruene Paletten im Lager zaehlen
   // Nur belegte Lagerplaetze beruecksichtigen.
   // 'Fehler' und 'Unbekannt' werden nicht mitgezaehlt.
   // =====================================================
   REGION Paletten nach Farbe zaehlen
       #Anzahl_Blau := 0;
       #Anzahl_Gruen := 0;
       #Anzahl_Unbekannte_Farbe := 0;
       FOR #i := 1 TO 54 DO

           IF NOT "HochregallagerDB".Lagerplaetze[#i].Frei THEN

               IF "HochregallagerDB".Lagerplaetze[#i].Materialfarbe S_COMP 'Blau' THEN
                   #Anzahl_Blau := #Anzahl_Blau + 1;

               ELSIF "HochregallagerDB".Lagerplaetze[#i].Materialfarbe S_COMP 'Gruen' THEN
                   #Anzahl_Gruen := #Anzahl_Gruen + 1;

               ELSIF "HochregallagerDB".Lagerplaetze[#i].Materialfarbe S_COMP 'Fehler' OR
                     "HochregallagerDB".Lagerplaetze[#i].Materialfarbe S_COMP 'Unbekannt'THEN
                   #Anzahl_Unbekannte_Farbe := #Anzahl_Unbekannte_Farbe + 1;
               END_IF;

           END_IF;

       END_FOR;
   END_REGION

   // =====================================================
   // 4. Palettendaten freier Lagerplaetze zuruecksetzen
   // Farbtext, Farbcode und Zeitstempel loeschen,
   // wenn der jeweilige Lagerplatz frei ist. 
   // =====================================================
   REGION Freie Lagerplaetze bereinigen

       FOR #i := 1 TO 54 DO

           // Palettendaten loeschen, wenn der Lagerplatz frei ist
           IF "HochregallagerDB".Lagerplaetze[#i].Frei THEN

               "HochregallagerDB".Lagerplaetze[#i].Materialfarbe := '';

               "HochregallagerDB".Lagerplaetze[#i].Materialfarbe_Nummer := 0;

               "HochregallagerDB".Lagerplaetze[#i].DatumUhrzeit :=
               DT#1990-01-01-00:00:00;

           END_IF;

       END_FOR;

   END_REGION

   // =====================================================
   // 5. Freie Lagerplaetze zaehlen und Lagerstatus auswerten
   // =====================================================
   // Anzahl der freien Lagerplaetze ermitteln
   REGION Lagerstatus und Warnungen

       #Anzahl_Freie_Plaetze := 0;

       FOR #i := 1 TO 54 DO
           IF "HochregallagerDB".Lagerplaetze[#i].Frei THEN
               #Anzahl_Freie_Plaetze := #Anzahl_Freie_Plaetze + 1;
           END_IF;
       END_FOR;

       // Warnung bei wenigen freien Lagerplaetzen, auch bei vollem Lager
       #Warnung_Wenig_Freie_Plaetze := #Anzahl_Freie_Plaetze <= #Warnschwelle_Freie_Plaetze;

       // Lager voll: Keine freien Lagerplaetze vorhanden
       #Lager_Voll := (#Anzahl_Freie_Plaetze = 0);


       // Sammelwarnung entsprechend dem aktuellen Lagerstatus aktualisieren
       #Warnung := #Warnung_Wenig_Freie_Plaetze OR #Lager_Voll;


       // Lager voll
       IF #Lager_Voll THEN
           #Warnung_Wenig_Freie_Plaetze := FALSE;
       END_IF;
   END_REGION
END_FUNCTION_BLOCK

FUNCTION_BLOCK "FB_ControlPanel"   // FB10, FBD
{ S7_Optimized_Access := 'FALSE' }
VERSION : 0.1
   VAR_INPUT
      IN_MS : Bool;   // Hauptschalter
      IN_ES : Bool;   // Not-Halt
      IN_Start : Bool;   // Start
      IN_Stop : Bool;   // Stop
      IN_FIO_RUN : Bool;   // Factory IO RUN
      IN_BLUE : Int;   // Blaue Teile
      IN_GREEN : Int;   // Grüne Teile
      IN_SIM : Bool;   // Stacker in Motion
      IN_CIM : Bool;   // Conveyor in Motion
      IN_ERROR : Bool;   // Störung
      IN_WARNING : Bool;   // Warnung
      IN_TT : Bool;   // Taktmerker
   END_VAR
   VAR_OUTPUT
      OUT_MSR : Bool;   // Meldesäule Rot
      OUT_MSY : Bool;   // Meldesäule Gelb
      OUT_MSG : Bool;   // Meldesäule Grün
      OUT_MLG : Bool;   // Anzeige Taster grün
      OUT_MLR : Bool;   // Anzeige Taster Rot
      OUT_RB : Bool;   // Rundumleuchte
      OUT_HORN : Bool;   // Sirene
      OUT_ESIO : Bool;   // Not-Halt IO
      OUT_GREEN : Int;   // Anzeige grüne Teile
      OUT_BLUE : Int;   // Anzeige Grüne Teile
      OUT_ME : Bool;   // Freigabe Bewegung
      OUT_SEOC : Bool;   // Stop Ende Zyklus
   END_VAR
   VAR
      "Not-Halt_IO" : Bool;   // Not-Halt in Ordnung
      Anlage_EIN : Bool;   // Anlage ist eingeschaltet
      Anlage_Warnung : Bool;   // Anlage Warnung
      Anlage_Störung : Bool;   // Anlage Störung
      Anlage_Start : Bool;   // Anlage gestartet
      Flanke_Start : Bool;   // Flanke Starttaster
      Anforderung_Stop : Bool;   // Anforderung Anlage Stop
      Flanke_Stop : Bool;   // Flanke Stoptaster
      Anlage_Stop : Bool;   // Anlage gestoppt
      Anlage_in_Bewegung : Bool;   // Anlage in Bewegung
      Betriebsbereit : Bool;   // Anlage Betriebsbereit
      In_Betrieb : Bool;   // Anlage in Betrieb
      Anlauf : Bool;   // Anlage im Anlauf
      Timer_Anlauf : TP;   // Timer Anlauf (10 Sek)
      Flanke_Anlauf : Bool;   // Flanke Anlauf beendet
      Flanke_Stillstand : Bool;
   END_VAR
   VAR_TEMP   // added for the SCL form of the ladder/FBD networks
      _w1 : Bool;
      _w2 : Bool;
      _w3 : Bool;
   END_VAR
BEGIN

REGION Network 1: Not-Halt
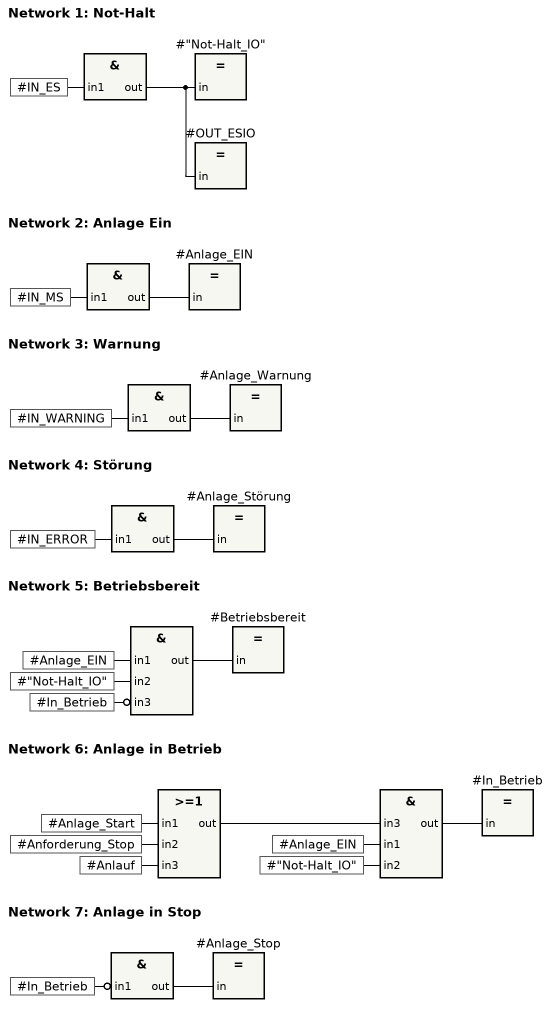
   #"Not-Halt_IO" := #IN_ES;
   #OUT_ESIO := #IN_ES;
END_REGION

REGION Network 2: Anlage Ein
   #Anlage_EIN := #IN_MS;
END_REGION

REGION Network 3: Warnung
   #Anlage_Warnung := #IN_WARNING;
END_REGION

REGION Network 4: Störung
   #Anlage_Störung := #IN_ERROR;
END_REGION

REGION Network 5: Betriebsbereit
   #Betriebsbereit := #Anlage_EIN AND #"Not-Halt_IO" AND NOT #In_Betrieb;
END_REGION

REGION Network 6: Anlage in Betrieb
   #In_Betrieb := (#Anlage_Start OR #Anforderung_Stop OR #Anlauf) AND #Anlage_EIN AND #"Not-Halt_IO";
END_REGION

REGION Network 7: Anlage in Stop
   #Anlage_Stop := NOT #In_Betrieb;
END_REGION

REGION Network 8: Anlauf
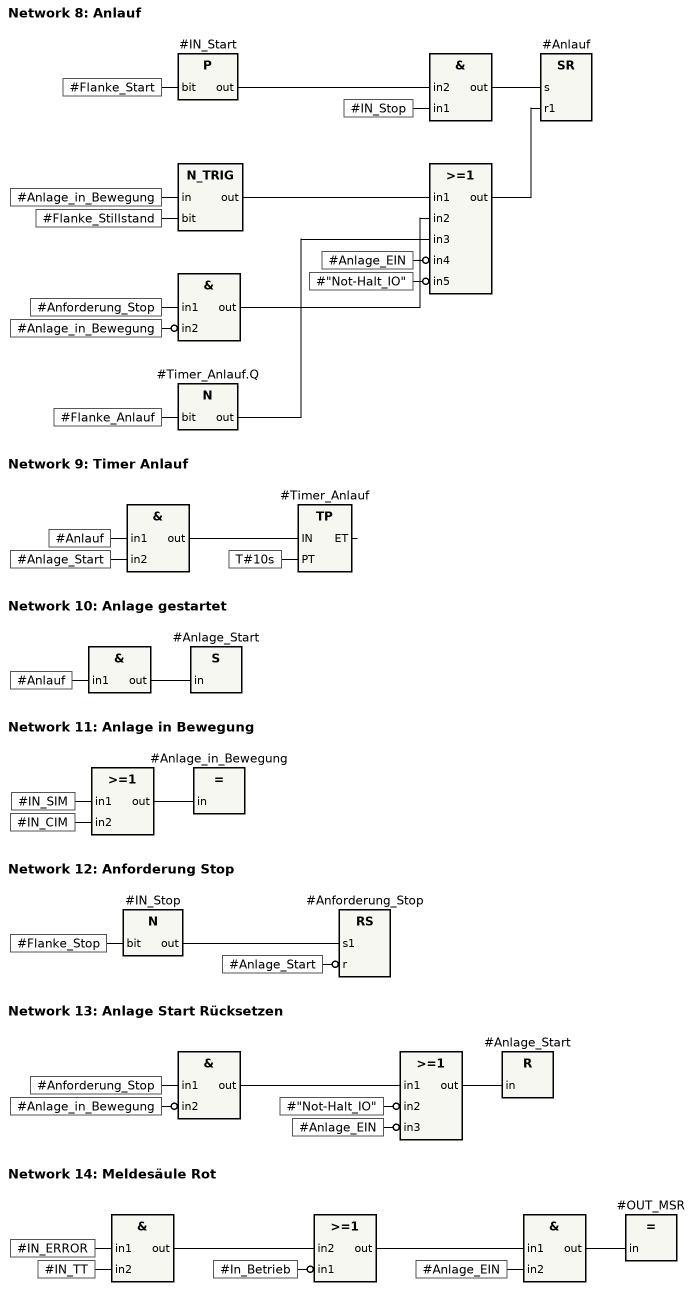
   #_w1 := #IN_Start AND NOT #Flanke_Start;   // rising edge of #IN_Start
   #Flanke_Start := #IN_Start;
   #_w2 := NOT #Anlage_in_Bewegung AND #Flanke_Stillstand;   // falling edge
   #Flanke_Stillstand := #Anlage_in_Bewegung;
   #_w3 := NOT #Timer_Anlauf.Q AND #Flanke_Anlauf;   // falling edge of #Timer_Anlauf.Q
   #Flanke_Anlauf := #Timer_Anlauf.Q;
   IF #_w1 AND #IN_Stop THEN
       #Anlauf := TRUE;   // SR flip-flop
   END_IF;
   IF #_w2 OR (#Anforderung_Stop AND NOT #Anlage_in_Bewegung) OR #_w3 OR NOT #Anlage_EIN OR NOT #"Not-Halt_IO" THEN
       #Anlauf := FALSE;
   END_IF;
END_REGION

REGION Network 9: Timer Anlauf
   #Timer_Anlauf.TP(IN := #Anlauf AND #Anlage_Start, PT := T#10s);
END_REGION

REGION Network 10: Anlage gestartet
   IF #Anlauf THEN #Anlage_Start := TRUE; END_IF;
END_REGION

REGION Network 11: Anlage in Bewegung
   #Anlage_in_Bewegung := #IN_SIM OR #IN_CIM;
END_REGION

REGION Network 12: Anforderung Stop
   #_w1 := NOT #IN_Stop AND #Flanke_Stop;   // falling edge of #IN_Stop
   #Flanke_Stop := #IN_Stop;
   IF NOT #Anlage_Start THEN
       #Anforderung_Stop := FALSE;   // RS flip-flop
   END_IF;
   IF #_w1 THEN #Anforderung_Stop := TRUE; END_IF;
END_REGION

REGION Network 13: Anlage Start Rücksetzen
   IF (#Anforderung_Stop AND NOT #Anlage_in_Bewegung) OR NOT #"Not-Halt_IO" OR NOT #Anlage_EIN THEN
       #Anlage_Start := FALSE;
   END_IF;
END_REGION

REGION Network 14: Meldesäule Rot
   #OUT_MSR := ((#IN_ERROR AND #IN_TT) OR NOT #In_Betrieb) AND #Anlage_EIN;
END_REGION

REGION Network 15: Meldesäule Gelb
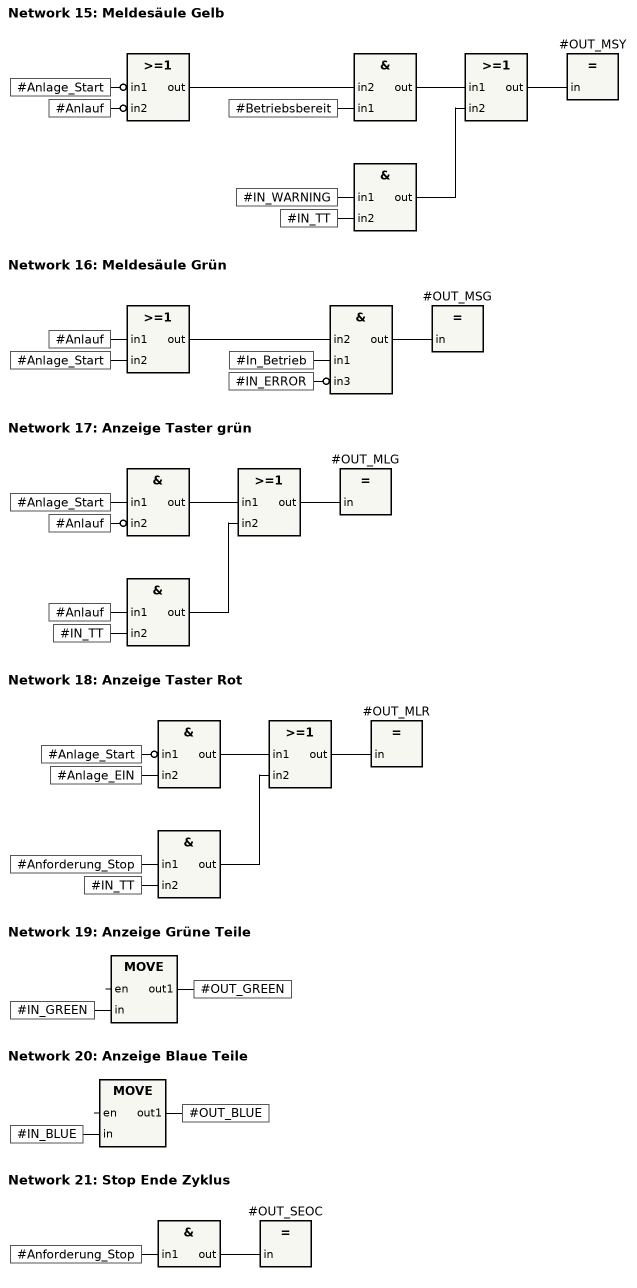
   #OUT_MSY := ((NOT #Anlage_Start OR NOT #Anlauf) AND #Betriebsbereit) OR (#IN_WARNING AND #IN_TT);
END_REGION

REGION Network 16: Meldesäule Grün
   #OUT_MSG := (#Anlauf OR #Anlage_Start) AND #In_Betrieb AND NOT #IN_ERROR;
END_REGION

REGION Network 17: Anzeige Taster grün
   #OUT_MLG := (#Anlage_Start AND NOT #Anlauf) OR (#Anlauf AND #IN_TT);
END_REGION

REGION Network 18: Anzeige Taster Rot
   #OUT_MLR := (NOT #Anlage_Start AND #Anlage_EIN) OR (#Anforderung_Stop AND #IN_TT);
END_REGION

REGION Network 19: Anzeige Grüne Teile
   #OUT_GREEN := #IN_GREEN;
END_REGION

REGION Network 20: Anzeige Blaue Teile
   #OUT_BLUE := #IN_BLUE;
END_REGION

REGION Network 21: Stop Ende Zyklus
   #OUT_SEOC := #Anforderung_Stop;
END_REGION

REGION Network 22: Freigabe Bewegung
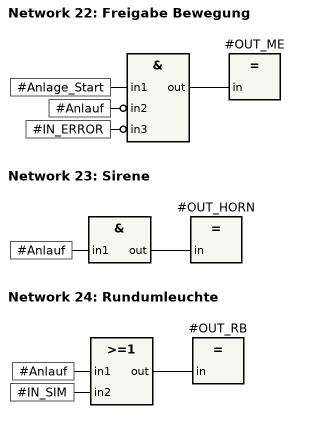
   #OUT_ME := #Anlage_Start AND NOT #Anlauf AND NOT #IN_ERROR;
END_REGION

REGION Network 23: Sirene
   #OUT_HORN := #Anlauf;
END_REGION

REGION Network 24: Rundumleuchte
   #OUT_RB := #Anlauf OR #IN_SIM;
END_REGION
END_FUNCTION_BLOCK

// folder: LAGER/FC

FUNCTION "FC_HMI_Bewegung" : Void   // FC1, SCL
{ S7_Optimized_Access := 'FALSE' }
VERSION : 0.1
   VAR_INPUT
      Position : Int;   // Ziellagerplatz fuer die HMI-Animation (1–54).
      Takt_Impuls : Bool;   // Taktsignal fuer die schrittweise Bewegung zum Ziel.
      Reset_Bewegung : Bool;   // Setzt die Bewegungszaehler bei deren Aufruf auf 0 zurueck.
   END_VAR
   VAR_OUTPUT
      HMI_X_Bewegung : Int;   // Aktueller horizontaler Verschiebungswert der HMI-Animation in Pixeln.
      HMI_Z_Bewegung : Int;   // Aktueller vertikaler Verschiebungswert der HMI-Animation in Pixeln.
   END_VAR
   VAR_TEMP
      Zeile : Int;   // Berechnete Zeile des Ziellagerplatzes (1–6).
      Spalte : Int;   // Berechnete Spalte des Ziellagerplatzes (1–9).
      X_Ziel : Int;   // Absolute horizontale Zielkoordinate in Pixeln.
      Y_Ziel : Int;   // Absolute vertikale Zielkoordinate in Pixeln.
      HMI_X_Ziel : Int;   // Horizontale Zielverschiebung relativ zur Referenz X = 120.
      HMI_Z_Ziel : Int;   // Vertikale Zielverschiebung relativ zur Referenz Y = 221.
      X_Counter_Ziel : Int;   // Zielzaehlerstand fuer X; ein Zaehlschritt entspricht 5 Pixeln.
      Z_Counter_Ziel : Int;   // Zielzaehlerstand fuer Z; ein Zaehlschritt entspricht 5 Pixeln.
   END_VAR
BEGIN
   // ---------------------------------------------------------
   // Zielposition berechnen
   // ---------------------------------------------------------
   IF (#Position >= 1) AND (#Position <= 54) THEN

       #Zeile := ((#Position - 1) / 9) + 1;
       #Spalte := ((#Position - 1) MOD 9) + 1;

       #X_Ziel := 175 + ((#Spalte - 1) * 62);
       #Y_Ziel := 172 - ((#Zeile - 1) * 51);

       #HMI_X_Ziel := #X_Ziel - 120;
       #HMI_Z_Ziel := #Y_Ziel - 221;
   ELSE
       #HMI_X_Bewegung := 1;
       #HMI_Z_Bewegung := 1;
       RETURN;
   END_IF;

   // ---------------------------------------------------------
   // Skalierte Zielwerte
   // 1 Counter-Schritt = 5 Pixel
   // ---------------------------------------------------------
   #X_Counter_Ziel := #HMI_X_Ziel / 5;
   #Z_Counter_Ziel := #HMI_Z_Ziel / 5;

   // ---------------------------------------------------------
   // CTUD X
   // ---------------------------------------------------------
   "IEC_Counter_x_DB".CTUD(
   CU := #Takt_Impuls AND
   ("IEC_Counter_x_DB".CV < #X_Counter_Ziel),

   CD := #Takt_Impuls AND
   ("IEC_Counter_x_DB".CV > #X_Counter_Ziel),

   R  := #Reset_Bewegung,
   LD := FALSE,

   PV := #X_Counter_Ziel
   );


   // Counterwert zurück in Pixel umrechnen
   #HMI_X_Bewegung := "IEC_Counter_x_DB".CV * 5;


   // ---------------------------------------------------------
   // CTUD Z
   // ---------------------------------------------------------

   "IEC_Counter_z_DB".CTUD(
                           CU := #Takt_Impuls AND
                           ("IEC_Counter_z_DB".CV < #Z_Counter_Ziel),

                           CD := #Takt_Impuls AND
                           ("IEC_Counter_z_DB".CV > #Z_Counter_Ziel),

                           R := #Reset_Bewegung,
                           LD := FALSE,

                           PV := #Z_Counter_Ziel
   );


   // Counterwert zurück in Pixel umrechnen
   #HMI_Z_Bewegung := "IEC_Counter_z_DB".CV * 5;
END_FUNCTION

FUNCTION "FC_Eingaben" : Void   // FC2, FBD
{ S7_Optimized_Access := 'FALSE' }
VERSION : 0.1
BEGIN

REGION Network 1: Hauptschalter 0-Aus, 1-Ein
END_REGION
END_FUNCTION

// folder: LAGER/Lager_AWL

FUNCTION "Lager_DB_löschen" : Void   // FC100, STL
{ S7_Optimized_Access := 'FALSE' }
VERSION : 0.1
// Mit diesem Baustein weden alle Datenworte des DB8000 gelöscht. Bei "löschen" = 1 wird der DB8000 Inhalt gelöscht.
   VAR_INPUT
      löschen : Bool;
   END_VAR
   VAR_OUTPUT
      Löschen_fertig : Bool;
   END_VAR
   VAR_TEMP
      HM_Schleifenzähler : DInt;
      HM_ADR : DWord;
      HM_Byte_Adr : DInt;
   END_VAR
BEGIN

REGION Network 1
         OPN   "Lager_Daten";

         A     #löschen;
         R     #Löschen_fertig;
         JCN   nix;


         L     DINT#54;

   SCHL: T     #HM_Schleifenzähler;

         L     #HM_Schleifenzähler;  // Bildung der speicherindirekten Adresse
         L     DINT#1;  // ( Schleifenzähler - 1 ) * 2 = Bytenummer
         -D;  //
         L     DINT#2;
         *D;
         T     #HM_Byte_Adr;

         SLD   3;  // Erzeugung der Bit-Adresse 0 = 0 durch schieben von 3 Stellen im DWORD (AKKU 1)
         T     #HM_ADR;  //  Bildung der indirekten Adresse

         L     0;
         T     DBW [ #HM_ADR];  // Beladen des Datenwortes mit 0

         L     #HM_Schleifenzähler;
         LOOP  SCHL;  // Wenn der #Schleifenzähler <= 0 wird die Schleife verlassen

         S     #Löschen_fertig;
   nix:  NOP   0;
END_REGION
END_FUNCTION

FUNCTION "Suche_Leeres_Fach" : Void   // FC101, STL
{ S7_Optimized_Access := 'FALSE' }
VERSION : 0.1
// Der Baustein dient zum Suchen einer Lagerfachnummer (1...54) mit den Werten  "1" für ein blaues Teil.
// Wird ein Fach gefunden beginnend vom Fach 1, so wird die Fachnummer ausgegeben. 
// Ist die Suche erfolglos, wird  Fachnummer = 0 und "Lager voll" = 1.  
// Mit dem Starteingang erfolgt die Ausführung.
// 
// Die Schnittstellenparameter "Lagerfach_Nr" und "Teil_nicht_vorhanden" sind als InOut-Parameter organisiert. Diese müssen mit Operanden, dessen  Daten über den AG-Zyklus hinaus erhalten bleiben. ( Merker, Datenbaustein-Daten , FB-Instanzen => Stat- Parameter)
// Der FC hat hierfür intern keine Möglichkeit.
   VAR_INPUT
      Start : Bool;
   END_VAR
   VAR_IN_OUT
      Lagerfach_Nr : Int;
      Lager_voll : Bool;
   END_VAR
   VAR_TEMP
      HM_Schleifenzähler : DInt;
      HM_Lagerfach_Nr : DInt;
   END_VAR
BEGIN

REGION Network 1
         A     #Start;
         JCN   ENDE;  // Ist Start = 0 überspringen aller Befehle

         OPN   "Lager_Daten";  // DB 8000 öffnen

         L     0;
         T     #HM_Lagerfach_Nr;  // Laden des Wertes 0  auf einen temporären Zwischenspeicher

         LAR1  P#0.0;
   // laden der Anfangsadresse mit Hilfe einer Pointer-Konstanten ( Adresse 0.0 ) in das Adressregister AR1
   // der CPU für die Adressregister indirekte Adressierung

         L     54;  // laden des Startwertes für die Loop-Schleife
   // Ziel ist es vom Lagerfach 1 beginnend zu suchen. Aus diesem Gund beginnt man mit dem Wert 54 ( höchste Fachnummer )
   // für den Schleifenzähler
   // Der Loop-Befehl verringert den AKKU1-Inhalt automatisch um 1.

   SCHL: T     #HM_Schleifenzähler;

         L     DBW [ AR1 , P#0.0 ];  // Laden des DBW mit der Anfangsadresse AR1 => 0.0 und einem Veratz von 0.0 => Resultat Adresse 0.0
         L     0;
         ==I;  // Untersuchung auf Inhalt = 0 für leeres Fach
         JCN   neu;  // Ist das nicht der Fall wird weiter gesucht
         L     55;  // Ermittelung der Fachnummer aus Subtraktion => Startwert = Max. Wert +1 ,
         L     #HM_Schleifenzähler;  // damit bei Adresse 0.0 die Fachnummer 1 ausgegeben wird.
         -I;
         T     #HM_Lagerfach_Nr;
         JU    POS;  // Ist ein Fach gefunden, wird die Suche beendet.
   neu:  +AR1  P#2.0;  // Sonst wird die im Adressregister AR1 vorhandene Adresse um 2 Byte
         NOP   0;  // für die Auswahl die nächste Fachuntersuchung (2.0) erhöht.

         L     #HM_Schleifenzähler;  // Vor dem Loop-Befehl wird der Speicher für den Schleifenzähler in den AKKU1 geladen.
         LOOP  SCHL;

         L     #HM_Lagerfach_Nr;  // Erzeugung der Meldung "Lager voll".
         L     0;
         ==I;
         =     #Lager_voll;
         JCN   ENDE;
         L     0;  // Bei "Lager voll" wird die Lagerfach-Nr.= 0 ausgeben.
         T     #Lagerfach_Nr;
         JU    ENDE;
   POS:  R     #Lager_voll;
         L     #HM_Lagerfach_Nr;
         T     #Lagerfach_Nr;
   ENDE: NOP   0;
END_REGION
END_FUNCTION

FUNCTION "Suche_Blau" : Void   // FC102, STL
{ S7_Optimized_Access := 'FALSE' }
VERSION : 0.1
// Der Baustein dient zum Suchen einer Lagerfachnummer (1...54) mit den Werten  "1" für Fach mit blauen Teil.
// Wird ein Fach gefunden beginnend vom Fach 1, so wird die Fachnummer ausgegeben. 
// Ist die Suche erfolglos, wird  Fachnummer = 0 und "kein_Teil_vorhanden" = 1 ausgegeben.  
// Mit dem Starteingang erfolgt die Ausführung.
// 
// Die Schnittstellenparameter "Lagerfach_Nr" und "kein Teil vorhanden" sind als InOut-Parameter organisiert. Diese müssen mit Operanden, dessen  Daten über den AG-Zyklus hinaus erhalten bleiben. 
// ( Merker, Datenbaustein-Daten , FB-Instanzen => Stat- Parameter)
// Der FC hat hierfür intern keine Möglichkeit.
   VAR_INPUT
      Start : Bool;
   END_VAR
   VAR_IN_OUT
      Lagerfach_Nr : Int;
      kein_Teil_vorhanden : Bool;
   END_VAR
   VAR_TEMP
      HM_Schleifenzähler : DInt;
      HM_Lagerfach_Nr : DInt;
   END_VAR
BEGIN

REGION Network 1
         A     #Start;
         JCN   ENDE;  // Ist Start = 0 überspringen aller Befehle

         OPN   "Lager_Daten";  // DB 8000 öffnen

         L     0;
         T     #HM_Lagerfach_Nr;  // Laden des Wertes 0  auf einen temporären Zwischenspeicher

         LAR1  P#0.0;
   // laden der Anfangsadresse mit Hilfe einer Pointer-Konstanten ( Adresse 0.0 ) in das Adressregister AR1
   // der CPU für die Adressregister indirekte Adressierung

         L     54;  // laden des Startwertes für die Loop-Schleife
   // Ziel ist es vom Lagerfach 1 beginnend zu suchen. Aus diesem Gund beginnt man mit dem Wert 54 ( höchste Fachnummer )
   // für den Schleifenzähler
   // Der Loop-Befehl verringert den AKKU1-Inhalt automatisch um 1.

   SCHL: T     #HM_Schleifenzähler;

         L     DBW [ AR1 , P#0.0 ];  // Laden des DBW mit der Anfangsadresse AR1 => 0.0 und einem Veratz von 0.0 => Resultat Adresse 0.0
         L     1;
         ==I;  // Untersuchung auf Inhalt = 1 für ein Fach mit blauen Teil
         JCN   neu;  // Ist das nicht der Fall wird weiter gesucht
         L     55;  // Ermittelung der Fachnummer aus Subtraktion => Startwert = Max. Wert +1 ,
         L     #HM_Schleifenzähler;  // damit bei Adresse 0.0 die Fachnummer 1 ausgegeben wird.
         -I;
         T     #HM_Lagerfach_Nr;
         JU    POS;  // Ist ein Fach gefunden, wird die Suche beendet.
   neu:  +AR1  P#2.0;  // Sonst wird die im Adressregister AR1 vorhandene Adresse um 2 Byte
         NOP   0;  // für die Auswahl die nächste Fachuntersuchung (2.0) erhöht.

         L     #HM_Schleifenzähler;  // Vor dem Loop-Befehl wird der Speicher für den Schleifenzähler in den AKKU1 geladen.
         LOOP  SCHL;

         L     #HM_Lagerfach_Nr;  // Erzeugung der Meldung "Teil nicht vorhanden".
         L     0;
         ==I;
         =     #kein_Teil_vorhanden;
         JCN   ENDE;
         L     0;  // Bei "kein Teil vorhanden" wird die Lagerfach-Nr.= 0 ausgeben.
         T     #Lagerfach_Nr;
         JU    ENDE;
   POS:  R     #kein_Teil_vorhanden;
         L     #HM_Lagerfach_Nr;
         T     #Lagerfach_Nr;
   ENDE: NOP   0;
END_REGION
END_FUNCTION

FUNCTION "Suche_Grün" : Void   // FC103, STL
{ S7_Optimized_Access := 'FALSE' }
VERSION : 0.1
// Der Baustein dient zum Suchen einer Lagerfachnummer (1...54) mit den Werten  "2" für ein grünes Teil im Fach.
// Wird ein Fach gefunden beginnend vom Fach 1, so wird die Fachnummer ausgegeben. 
// Ist die Suche erfolglos, wird  Fachnummer = 0 und "kein Teil vorhanden" = 1 ausgegeben.  
// Mit dem Starteingang erfolgt die Ausführung.
// 
// Die Schnittstellenparameter "Lagerfach_Nr" und "Lager voll" sind als InOut-Parameter organisiert. Diese müssen mit Operanden, dessen  Daten über den AG-Zyklus hinaus erhalten bleiben. 
// ( Merker, Datenbaustein-Daten , FB-Instanzen => Stat- Parameter)
// Der FC hat hierfür intern keine Möglichkeit.
   VAR_INPUT
      Start : Bool;
   END_VAR
   VAR_IN_OUT
      Lagerfach_Nr : Int;
      kein_Teil_vorhanden : Bool;
   END_VAR
   VAR_TEMP
      HM_Schleifenzähler : DInt;
      HM_Lagerfach_Nr : DInt;
   END_VAR
BEGIN

REGION Network 1
         A     #Start;
         JCN   ENDE;  // Ist Start = 0 überspringen aller Befehle

         OPN   "Lager_Daten";  // DB 8000 öffnen

         L     0;
         T     #HM_Lagerfach_Nr;  // Laden des Wertes 0  auf einen temporären Zwischenspeicher

         LAR1  P#0.0;
   // laden der Anfangsadresse mit Hilfe einer Pointer-Konstanten ( Adresse 0.0 ) in das Adressregister AR1
   // der CPU für die Adressregister indirekte Adressierung

         L     54;  // laden des Startwertes für die Loop-Schleife
   // Ziel ist es vom Lagerfach 1 beginnend zu suchen. Aus diesem Gund beginnt man mit dem Wert 54 ( höchste Fachnummer )
   // für den Schleifenzähler
   // Der Loop-Befehl verringert den AKKU1-Inhalt automatisch um 1.

   SCHL: T     #HM_Schleifenzähler;

         L     DBW [ AR1 , P#0.0 ];  // Laden des DBW mit der Anfangsadresse AR1 => 0.0 und einem Veratz von 0.0 => Resultat Adresse 0.0
         L     2;
         ==I;  // Untersuchung auf Inhalt = 2 für ein Fach mit grünen Teil
         JCN   neu;  // Ist das nicht der Fall wird weiter gesucht
         L     55;  // Ermittelung der Fachnummer aus Subtraktion => Startwert = Max. Wert +1 ,
         L     #HM_Schleifenzähler;  // damit bei Adresse 0.0 die Fachnummer 1 ausgegeben wird.
         -I;
         T     #HM_Lagerfach_Nr;
         JU    POS;  // Ist ein Fach gefunden, wird die Suche beendet.
   neu:  +AR1  P#2.0;  // Sonst wird die im Adressregister AR1 vorhandene Adresse um 2 Byte
         NOP   0;  // für die Auswahl die nächste Fachuntersuchung (2.0) erhöht.

         L     #HM_Schleifenzähler;  // Vor dem Loop-Befehl wird der Speicher für den Schleifenzähler in den AKKU1 geladen.
         LOOP  SCHL;

         L     #HM_Lagerfach_Nr;  // Erzeugung der Meldung "Teil nicht vorhanden".
         L     0;
         ==I;
         =     #kein_Teil_vorhanden;
         JCN   ENDE;
         L     0;  // Bei "Teil nicht vorhanden" wird die Lagerfach-Nr.= 0 ausgeben.
         T     #Lagerfach_Nr;
         JU    ENDE;
   POS:  R     #kein_Teil_vorhanden;
         L     #HM_Lagerfach_Nr;
         T     #Lagerfach_Nr;
   ENDE: NOP   0;
END_REGION
END_FUNCTION

FUNCTION "Lagerfach_beschreiben" : Void   // FC104, STL
{ S7_Optimized_Access := 'FALSE' }
VERSION : 0.1
// Der Baustein dient zum Beschreiben einer Lagerfachnummer (1...54) mit den Werten  "1" für Belegung mit einem blauen Teil oder dem Wert  "2" für ein grünes Teil oder mit Wert "0" für ein leeres Fach.
// Das Beschreiben erfolgt durch Vorwahl der Lagerfachnummer und der Auswahl an den Eigängen für blau oder grün.
// Mit dem Starteingang erfolgt die Ausführung.
// Die Fehleranzeige wird dann aktiviert, wenn die Lagerfachnummer nicht im Bereich von 1..54 liegt  oder die Auswahlen nicht  oder mehrere aktiv sind.
// In diesem Fall bleibt das Lagerfach im DB8000 unverändert.
   VAR_INPUT
      Start : Bool;
      Blau : Bool;   // Blau = 1
      Grün : Bool;   // Grün = 2
      Leer : Bool;   // Leer = 0
      Lagerfach_Nr : Int;
   END_VAR
   VAR_OUTPUT
      Fehler : Bool;
   END_VAR
   VAR_TEMP
      HM_Schleifenzähler : DInt;
      HM_Lagerfach_Nr : DInt;
      HM_Adr : DWord;
   END_VAR
BEGIN

REGION Network 1

         A     #Start;
         R     #Fehler;  // Bei Start löschen des Fehlerausganges
         JCN   NIX;  // Ist Start = 0 überspringen aller Befehle

         OPN   "Lager_Daten";  // DB 8000 öffnen

         A(;  // Untersuchung der Lagerfachnummer (1..54) sonst Fehler
         L     #Lagerfach_Nr;
         L     1;
         >=I;
         );
         A(;
         L     #Lagerfach_Nr;
         L     54;
         <=I;
         );
         JCN   Fehl;

         A     #Blau;  // Untersuchung der gleichzeitigen Aktivierung von "Leer", "Blau" und "Grün"
         AN    #Grün;  // sonst Fehler
         AN    #Leer;  // Es darf nur 1 Auswahl erfolgen. Fehler auch bei keiner Auswahl
         O;
         AN    #Blau;
         A     #Grün;
         AN    #Leer;
         O;
         AN    #Blau;
         AN    #Grün;
         A     #Leer;
         JCN   Fehl;

         L     #Lagerfach_Nr;  // Bildung der Anfangsadresse für das Lagerfach
         L     1;  // ( Fachnummer - 1) *2 => Anfangsadresse (Byte-Nummer)
         -I;
         L     2;
         *I;
         SLD   3;  // Bildung der speicherindirekten Adresse [Byte-Nummer Bit-Nummer
         T     #HM_Adr;  // Die Bit-Nummer muß ab  Byte-Zugriff = 0 sein.
         NOP   0;  // ( Schieben nach links 3 Stellen im DWORD )

         A     #Blau;
         AN    #Grün;
         AN    #Leer;
         JCN   Blau;  // Auswahl Blau sonst überspringen der Befehlzeilen
         L     1;  // Wert 1 für Blau
         T     DBW [ #HM_Adr];  // Laden in des DBW x durch speicherindirekte Adressierung

         JU    NIX;  // gehe zu Marke NIX

   Blau: NOP   0;

         A     #Grün;
         AN    #Blau;
         AN    #Leer;
         JCN   Leer;  // Auswahl Grün sonst überspringen der Befehlzeilen
         L     2;  // Wert 2 für Grün
         T     DBW [ #HM_Adr];  // Laden in des DBW x durch speicherindirekte Adressierung

         JU    NIX;  // gehe zu Marke NIX

   Leer: NOP   0;
         AN    #Grün;
         AN    #Blau;
         A     #Leer;
         JCN   NIX;  // Auswahl Leer sonst überspringen der Befehlzeilen
         L     0;  // Wert 0 für Leer
         T     DBW [ #HM_Adr];  // Laden in des DBW x durch speicherindirekte Adressierung

         JU    NIX;  // gehe zu Marke NIX

   Fehl: S     #Fehler;  // Bei Fehler setzen des Ausganges

   NIX:  NOP   0;
END_REGION
END_FUNCTION

// folder: Versand

FUNCTION_BLOCK "621_Suche_neu"   // FB5, SCL
{ S7_Optimized_Access := 'FALSE' }
VERSION : 0.1
   VAR_INPUT
      Betriebsbereit : Bool;
      "I_Taster GN" : Bool;
      "I_Taster BL" : Bool;
      I_Ausgelagert : Bool;
      I_Kontrolliert : Bool;
      I_Fehler : Bool;
   END_VAR
   VAR_OUTPUT
      Q_LED_GN : Bool;
      Q_LED_BL : Bool;
      Anforderung : Bool;
   END_VAR
   VAR_IN_OUT
      Lagerplaetze : Array[1..54] of "Datenspeicher";   // Lagerdaten der 54 Lagerplätze: Belegung, Farbe und Einlagerungszeit
      Fachnummer : Int;
      Farbcode : Int;
   END_VAR
   VAR
      s_suchfarbcode : Int;
      s_datum : Date_And_Time;
   END_VAR
   VAR_TEMP
      idx : Int;
   END_VAR
BEGIN
   IF NOT #Betriebsbereit THEN
       #Q_LED_GN := 0;
       #Q_LED_BL := 0;
       #Anforderung := 0;
       #Fachnummer := 0;
       #Farbcode := 0;
       #s_suchfarbcode := 0;
       #Q_LED_GN := 0;
       #Q_LED_BL := 0;
   ELSE
       IF #"I_Taster GN" AND NOT (#s_suchfarbcode = 1) THEN
           #s_suchfarbcode := 2;
       END_IF;
       IF #"I_Taster BL" AND  NOT (#s_suchfarbcode = 2) THEN
           #s_suchfarbcode := 1;
       END_IF;
       IF #I_Kontrolliert THEN
           #s_suchfarbcode := 0;
           #Farbcode := 0;
           #Anforderung := 0;
       END_IF;


       IF #s_suchfarbcode > 0 AND #Farbcode = 0 AND NOT #I_Kontrolliert THEN
           #Fachnummer := 0;
           FOR #idx := 1 TO 54 DO
               IF #Lagerplaetze[#idx].Materialfarbe_Nummer = #s_suchfarbcode AND (#Fachnummer = 0 OR #s_datum T_COMP #Lagerplaetze[#idx].DatumUhrzeit) THEN
                   #Fachnummer := #idx;
                   #s_datum := #Lagerplaetze[#idx].DatumUhrzeit;
                   #Farbcode := #s_suchfarbcode;
                   #Anforderung := 1;
               END_IF;
           END_FOR;
       END_IF;


       #Q_LED_GN := ((#s_suchfarbcode = 0) AND "Takt_1HZ") OR ((#Farbcode = 2) AND (#Fachnummer > 0));
       #Q_LED_BL := ((#s_suchfarbcode = 0) AND NOT "Takt_1HZ") OR ((#Farbcode = 1) AND (#Fachnummer > 0));
   END_IF;
END_FUNCTION_BLOCK

FUNCTION_BLOCK "609_DB zürücksetzen"   // FB6, SCL
{ S7_Optimized_Access := 'FALSE' }
VERSION : 0.1
   VAR_INPUT
      reset : Bool;
   END_VAR
   VAR_TEMP
      idx : Int;
   END_VAR
BEGIN
   IF #reset THEN
       FOR #idx := 1 TO 54 DO
           "HochregallagerDB".Lagerplaetze[#idx].Frei := 1;
       END_FOR;
   END_IF;
END_FUNCTION_BLOCK

FUNCTION_BLOCK "600_Versand_Main"   // FB600, FBD
{ S7_Optimized_Access := 'FALSE' }
AUTHOR : DJonas
VERSION : 0.1
   VAR_INPUT
      Start : Bool;
      Stop : Bool;
      "In Betrieb" : Bool;
      NotHalt : Bool;
   END_VAR
   VAR_IN_OUT
      Pult_Daten : "Datenaustausch_Versand";
   END_VAR
   VAR
      Ware_Holen : Bool;
      t_übergabe : Bool;
      t_kontrolliert : Bool;
      t_630Work : Bool;
      t_startrb : Bool;
      t_anforderung : Bool;
      t_ausgelagert : Bool;
      t_fehler : Bool;
      t_rbfrei : Bool;
      t_630_Grundstellung : Bool;
      s_ptrig : Bool;
      t_farbsensor : Int;
      t_fach : Int;
      t_farbe : Int;
      t_fachnummer : Int;
      t_farbcode : Int;
      "621_Suche_neu_Instance" : "621_Suche_neu";
      "630_Lagerfach holen_Instance_1" : "630_Lagerfach holen";
      "640_Rollenbahnen_Instance" : "640_Rollenbahnen";
      "609_DB zürücksetzen_Instance" : "609_DB zürücksetzen";
      IEC_Timer_0_Instance : TON;
   END_VAR
   VAR_TEMP
      t_630_atwork : Bool;
      t_safe : Bool;
   END_VAR
   VAR_TEMP   // added for the SCL form of the ladder/FBD networks
      _w1 : Bool;
   END_VAR
BEGIN

REGION Network 1
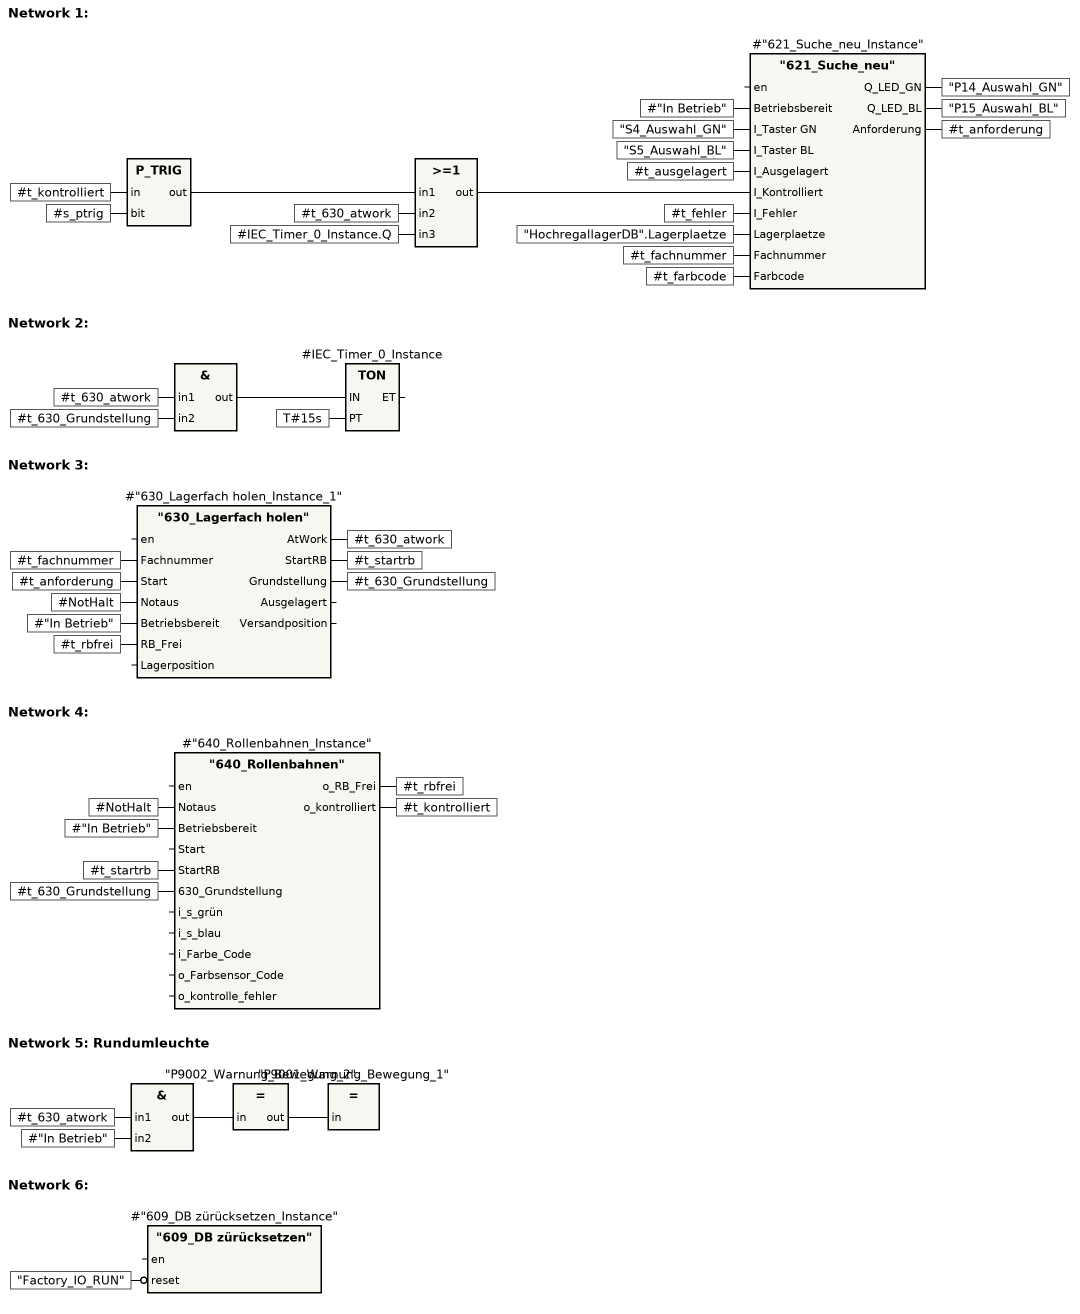
   #_w1 := #t_kontrolliert AND NOT #s_ptrig;   // rising edge
   #s_ptrig := #t_kontrolliert;
   #"621_Suche_neu_Instance"(Betriebsbereit := #"In Betrieb",   // "621_Suche_neu"
                           "I_Taster GN" := "S4_Auswahl_GN",
                           "I_Taster BL" := "S5_Auswahl_BL",
                           I_Ausgelagert := #t_ausgelagert,
                           I_Kontrolliert := #_w1 OR #t_630_atwork OR #IEC_Timer_0_Instance.Q,
                           I_Fehler := #t_fehler,
                           Lagerplaetze := "HochregallagerDB".Lagerplaetze,
                           Fachnummer := #t_fachnummer,
                           Farbcode := #t_farbcode,
                           Q_LED_GN => "P14_Auswahl_GN",
                           Q_LED_BL => "P15_Auswahl_BL",
                           Anforderung => #t_anforderung);
END_REGION

REGION Network 2
   #IEC_Timer_0_Instance.TON(IN := #t_630_atwork AND #t_630_Grundstellung, PT := T#15s);
END_REGION

REGION Network 3
   #"630_Lagerfach holen_Instance_1"(Fachnummer := #t_fachnummer,   // "630_Lagerfach holen"
                           Start := #t_anforderung,
                           Notaus := #NotHalt,
                           Betriebsbereit := #"In Betrieb",
                           RB_Frei := #t_rbfrei,
                           AtWork => #t_630_atwork,
                           StartRB => #t_startrb,
                           Grundstellung => #t_630_Grundstellung);
END_REGION

REGION Network 4
   #"640_Rollenbahnen_Instance"(Notaus := #NotHalt,   // "640_Rollenbahnen"
                           Betriebsbereit := #"In Betrieb",
                           StartRB := #t_startrb,
                           "630_Grundstellung" := #t_630_Grundstellung,
                           o_RB_Frei => #t_rbfrei,
                           o_kontrolliert => #t_kontrolliert);
END_REGION

REGION Network 5: Rundumleuchte
   "P9002_Warnung_Bewegung_2" := #t_630_atwork AND #"In Betrieb";
   "P9001_Warnung_Bewegung_1" := "P9002_Warnung_Bewegung_2";
END_REGION

REGION Network 6
   #"609_DB zürücksetzen_Instance"(reset := NOT "Factory_IO_RUN");   // "609_DB zürücksetzen"
END_REGION
END_FUNCTION_BLOCK

FUNCTION_BLOCK "620_FB_Farbauswahl_Jewgeni_V2"   // FB620, SCL
{ S7_Optimized_Access := 'FALSE' }
AUTHOR : Jewgeni
VERSION : 0.1
   VAR_INPUT
      I_Taster_Gruen : Bool;
      I_Taster_Blau : Bool;
      I_Palette_Kontrolliert : Bool;
      I_Anlage_Aktiv : Bool;
      I_Farbsensor_Code : Int;
   END_VAR
   VAR_OUTPUT
      Q_LED_Gruen : Bool;
      Q_LED_Blau : Bool;
      Q_Fachnummer : Int;
      Q_Farbe_Code : Int;
      Q_Uebergabe_Aktiv : Bool;
      Q_Fehler_FalscheFarbe : Bool;
   END_VAR
   VAR_IN_OUT
      IQ_Lager_Regal : Array[1..54] of Int;
      O_GN : Int;
      O_BL : Int;
   END_VAR
   VAR
      stat_FP_Taster_Gruen : Bool;
      stat_Flanke_Gruen_Aktiv : Bool;
      stat_FP_Taster_Blau : Bool;
      stat_Flanke_Blau_Aktiv : Bool;
      stat_Schritt : Int;
      stat_GewaehlteFarbe : Int;
      stat_Fehler_FalscheFarbe : Bool;
   END_VAR
   VAR_TEMP
      idx : Int;
   END_VAR
BEGIN
   // SICHERHEIT: Wenn die Anlage stoppt (STOP / NOT-HALT), wird deine Auswahl sofort gelöscht
   IF NOT #I_Anlage_Aktiv THEN
       #stat_Schritt := 0;
       #Q_LED_Gruen := FALSE;
       #Q_LED_Blau := FALSE;
       #Q_Uebergabe_Aktiv := FALSE;
       #Q_Fachnummer := 0;
       #Q_Farbe_Code := 0;
       RETURN;
   END_IF;

   // --- S7-300 FLANKENAUSWERTUNG ---
   #stat_Flanke_Gruen_Aktiv := #I_Taster_Gruen AND NOT #stat_FP_Taster_Gruen;
   #stat_FP_Taster_Gruen := #I_Taster_Gruen;

   #stat_Flanke_Blau_Aktiv := #I_Taster_Blau AND NOT #stat_FP_Taster_Blau;
   #stat_FP_Taster_Blau := #I_Taster_Blau;


   // --- SCHRITTKETTE ---
   CASE #stat_Schritt OF

       0: // --- GRUNDSTELLUNG: Auf Auswahl durch den Bediener warten ---
           #Q_Uebergabe_Aktiv := FALSE;

           IF #stat_Flanke_Gruen_Aktiv THEN
               #stat_GewaehlteFarbe := 2; // 2 = Grün (Laut Projektvorgabe)
               #Q_LED_Gruen := TRUE;      // LED am Schaltkasten einschalten
               #stat_Schritt := 10;
           ELSIF #stat_Flanke_Blau_Aktiv THEN
               #stat_GewaehlteFarbe := 1; // 1 = Blau (Laut Projektvorgabe)
               #Q_LED_Blau := TRUE;       // LED am Schaltkasten einschalten
               #stat_Schritt := 10;
           END_IF;

       10: // --- SUCHE IM Übergebenen Array ---
           #Q_Fachnummer := 0;



          FOR #idx := 1 TO 54 DO
               // Greift jetzt absolut autark auf die Schnittstelle zu:
              IF #IQ_Lager_Regal[#idx] = #stat_GewaehlteFarbe THEN
                   #Q_Fachnummer := #idx;                 // Gefundene Fachnummer sichern
                   #Q_Farbe_Code := #stat_GewaehlteFarbe; // Farbcode mitsenden
                   EXIT;                                // Suche erfolgreich abbrechen
               END_IF;
           END_FOR;

           // Auswertung des Suchlaufs
           IF #Q_Fachnummer > 0 THEN
               #Q_Uebergabe_Aktiv := TRUE; // Belal signalisieren: "Fachnummer liegt an, du kannst holen!"
               #stat_Schritt := 20;        // Wechsel in den Wartemodus
           ELSE
               // Falls kein Teil dieser Farbe mehr im Lager ist: LEDs zurücksetzen, zurück auf Anfang
               #Q_LED_Gruen := FALSE;
               #Q_LED_Blau := FALSE;
               #stat_Schritt := 0;
           END_IF;

       20: // --- WARTEN AUF FERTIGMELDUNG & SENSORPRÜFUNG ---

           // 1. Fehlerprüfung: Wenn ein Teil am Sensor ist, muss die Farbe stimmen
           IF #I_Farbsensor_Code <> 0 THEN
               IF #I_Farbsensor_Code <> #stat_GewaehlteFarbe THEN
                   #Q_Fehler_FalscheFarbe := TRUE; // Alarm: Falsche Farbe gegriffen!
                   #Q_Uebergabe_Aktiv := FALSE;     // Folgesteuerung (Belal) sofort stoppen
               ELSE
                   #Q_Fehler_FalscheFarbe := FALSE; // Farbe ist korrekt
               END_IF;
           END_IF;

           // 2. Normaler Prozessabschluss (nur wenn kein Fehler ansteht)
           IF #I_Palette_Kontrolliert AND NOT #stat_Fehler_FalscheFarbe THEN
               #Q_LED_Gruen := FALSE;
               #Q_LED_Blau := FALSE;
               #Q_Uebergabe_Aktiv := FALSE;
               #stat_Schritt := 0; // Zurück in Grundstellung für nächsten Auftrag
           END_IF;

           // 3. Fehler-Quittierung (Manuell oder über Anlage_Aktiv-Reset)
           IF NOT #I_Anlage_Aktiv THEN
               #Q_Fehler_FalscheFarbe := FALSE; // Reset bei Anlagen-Stopp
           END_IF;

   END_CASE;
END_FUNCTION_BLOCK

FUNCTION_BLOCK "630_Lagerfach holen"   // FB630, SCL
{ S7_Optimized_Access := 'FALSE' }
AUTHOR : DJonas
VERSION : 0.1
   VAR_INPUT
      Fachnummer : Int;
      Start : Bool;
      Notaus : Bool;
      Betriebsbereit : Bool;
      RB_Frei : Bool;
      Lagerposition : Int;
   END_VAR
   VAR_OUTPUT
      AtWork : Bool;
      StartRB : Bool;
      Grundstellung : Bool;
      Ausgelagert : Bool;
      Versandposition : Int;
   END_VAR
   VAR
      "Wagen benutzt" : Bool;
      hilfsmerker_fahren : Bool;
      bewegung : Bool;
      Neutstart : Bool;
      Schritt : Int;
      Portal_Ist : Int;
      Portal_soll : Int;
      Schritt1Anlauf : TON;
      TON_Schritt11 : TON;
   END_VAR
BEGIN
       REGION Betriebsbereitschaft
           IF NOT #Notaus THEN
               #Schritt := 70;
               "STAPL_9001_Fachposition" := 0;
           ELSE
               IF #Schritt = 70 AND #Betriebsbereit THEN
                   "STAPL_9001_links_ausfahren" := 0;
                   "STAPL_9001_rechts_ausfahren" := 0;
                   #Neutstart := 1;
                   #Schritt := 8;
               END_IF;
           END_IF;

           #StartRB := 0;
           #Grundstellung := (#Schritt = 0) OR (#Schritt = 19);
           #AtWork := (#Schritt > 0 AND #Schritt < 70);

           #Schritt1Anlauf(IN := #AtWork, PT := T#1s);
           #TON_Schritt11(IN := #hilfsmerker_fahren, PT := T#2s);

           IF ( #Schritt = 0 AND NOT #Start) OR #Schritt = 70 THEN RETURN; END_IF;

       END_REGION
       REGION Bewegungsvariable
           #bewegung := "B9023_STAPL_Bew_X_aktiv"
           OR "B9024_STAPL_Bew_Z_aktiv"
           OR (NOT "B9020_STAPL_9001_Endlage_links" AND "STAPL_9001_links_ausfahren")
           OR (NOT "B9022_STAPL_9001_Endlage_rechts" AND "STAPL_9001_rechts_ausfahren")
           OR (NOT "B9021_STAPL_9001_Mittel_Pos" AND NOT "STAPL_9001_links_ausfahren" AND NOT "STAPL_9001_rechts_ausfahren");
       END_REGION
       REGION Start
           // Grundstellungsfahrt nacht Neustart/Nothalt einleiten
           IF #Betriebsbereit AND #Grundstellung = 0 AND #AtWork = 0 AND #Schritt = 70 THEN
               #AtWork := 1;
               #Schritt := 8;
           END_IF;

           // Fachabholung starten
           IF #Start AND #Schritt = 0 AND #Fachnummer > 0 THEN
               #Portal_Ist := "STAPL_9001_Fachposition";                   // Istposition zwischenspeichern
               #Portal_soll := #Fachnummer;                                // Sollposition zwischenspeichern
               IF #Portal_Ist = #Portal_soll OR #Portal_soll = 55 THEN     // Wenn Istposition gleich Sollposition oder Sollposition = 55
   //                "STAPL_9001_links_ausfahren" := 0;                      // Dann links ausfahren zurücksetzen (fals gesetzte) und zu Schritt 11 gehen
                   #Schritt := 11;
               ELSE                                                        // komplette schrittkette durchlaufen
                   #Portal_soll := #Portal_soll;
                   #Schritt := 1;
               END_IF;
           END_IF;
           // Warten bei Neustart
           IF NOT #Schritt1Anlauf.Q THEN
               RETURN;
           END_IF;

       END_REGION

       // Kollisionsverhinderung
       // wenn links ausfahren angesteuert, wird die fachnummer übergeben
       // 
       IF "STAPL_9001_links_ausfahren" THEN
           #Versandposition := #Portal_soll;
       END_IF;
       IF "B9021_STAPL_9001_Mittel_Pos" THEN
           #Versandposition := 0;
       END_IF;


   // Schrittkette
       CASE #Schritt OF
           1:  // von Grundstellung zu Fach fahren
               IF #bewegung THEN
                   #Schritt := 2;
               END_IF;
               IF #Portal_Ist = 55 OR #Portal_Ist = 0 THEN
                   "STAPL_9001_Fachposition" := #Portal_soll;
                   "STAPL_9001_Palette_heben" := 0;
               END_IF;
           2:  // nach links ausfahren
               IF NOT "B9020_STAPL_9001_Endlage_links" AND NOT #bewegung AND NOT ( #Lagerposition = #Portal_soll) THEN
                   "STAPL_9001_links_ausfahren" := 1;
                   #Schritt := 3;
               END_IF;
           3: // Palette anheben
               IF "B9020_STAPL_9001_Endlage_links" AND NOT #bewegung THEN
                   "STAPL_9001_Palette_heben" := 1;
                   IF #Fachnummer > 0 AND #Fachnummer < 55 THEN
                       "HochregallagerDB".Lagerplaetze[#Fachnummer].Frei := 1;
                   END_IF;
               END_IF;
               IF "STAPL_9001_Palette_heben" AND #bewegung THEN
                   #Schritt := 8;
               END_IF;
           8: // in Mittelstellung fahren und Startpunkt für Grundstellungsfahrt
               IF ("B9020_STAPL_9001_Endlage_links" OR "STAPL_9001_links_ausfahren") AND NOT #bewegung THEN
                   "STAPL_9001_links_ausfahren" := 0;
               END_IF;
               IF NOT "STAPL_9001_links_ausfahren" AND "B9021_STAPL_9001_Mittel_Pos" THEN
                   #Schritt := 9;
               END_IF;
           9: // Palette aus Fach nehmen abgeschlossen
               IF "B9021_STAPL_9001_Mittel_Pos" AND NOT #bewegung THEN
                   #Schritt := 11;
               END_IF;
           11: // zum Absetzen fahren
               IF #bewegung OR #TON_Schritt11.Q THEN
                   #Schritt := 15;
               END_IF;
               IF "B9021_STAPL_9001_Mittel_Pos" AND NOT #bewegung THEN
                   "STAPL_9001_Fachposition" := 55;
                   "STAPL_9001_Palette_heben" := 1;
                   #hilfsmerker_fahren := 1;
               END_IF;
           15: // Palette nach rechts fahren und senken
               IF #RB_Frei AND "STAPL_9001_Palette_heben" AND "B9021_STAPL_9001_Mittel_Pos" AND NOT #bewegung THEN
                   #hilfsmerker_fahren := 0;
                   "STAPL_9001_rechts_ausfahren" := 1;
               END_IF;
               IF "B9022_STAPL_9001_Endlage_rechts" AND "STAPL_9001_rechts_ausfahren" THEN
                   "STAPL_9001_Palette_heben" := 0;
                   #Schritt := 17;
               END_IF;
           17: // Palette senken
               IF NOT "STAPL_9001_Palette_heben" AND #bewegung THEN
                   #Schritt := 18;
               END_IF; 
           18: // in Mittelstellung fahren, Grundstellung erreicht
               IF NOT #bewegung THEN
                   "STAPL_9001_rechts_ausfahren" := 0;
                   #Schritt := 19;
               END_IF;
           19:
               IF "B9021_STAPL_9001_Mittel_Pos" AND NOT #Start THEN
                   #Schritt := 0;
                   IF #Neutstart THEN
                       #Neutstart := 0;
                   ELSE
                       #StartRB := 1;
                   END_IF;
               END_IF;
       END_CASE;
END_FUNCTION_BLOCK

